(* IEC 61131-3 sources: plc-st-coding-agent/progress/evidence/f14_v3_parallel_20261112/jobs/custom_minimax-m27 (part 3) *)

(* ---- self-hard-02.raw_candidate_01.st ---- *)
FUNCTION_BLOCK FB
VAR_INPUT
    startBtn   : BOOL;
    abortBtn   : BOOL;
    setpoint   : REAL;
    pv         : REAL;
    maxDuration: INT;
END_VAR
VAR_OUTPUT
    elapsed : INT := 0;
    phase   : INT := 0;
    timeout : BOOL := FALSE;
END_VAR
VAR
    prev_startBtn : BOOL := FALSE;
    prev_phase    : INT  := 0;
    risingEdge    : BOOL;
END_VAR

    // Detect rising edge of startBtn before any state changes this scan
    risingEdge := startBtn AND NOT prev_startBtn;

    // Priority 1: abort
    IF abortBtn THEN
        phase   := 9;
        // elapsed and timeout stay frozen (no assignment)

    // Priority 2: new rising edge (only if not aborted this scan)
    ELSIF risingEdge THEN
        elapsed := 0;
        timeout := FALSE;
        phase   := 1;

    // Priority 3: running phases — count and evaluate transition
    ELSIF (prev_phase = 1) OR (prev_phase = 2) THEN
        elapsed := elapsed + 1;

        // Check timeout before setting phase
        IF elapsed >= maxDuration THEN
            timeout := TRUE;
            phase   := 3;
        ELSE
            // Phase transition based on temperature
            IF (prev_phase = 2) OR (pv >= setpoint) THEN
                phase := 2;
            ELSE
                phase := 1;
            END_IF;
        END_IF;

    // Frozen states (phase 0, 3, 9) — no changes to elapsed/phase/timeout
    ELSE
        // phase, elapsed, timeout retain their values
    END_IF;

    // Update previous-cycle snapshot for next scan
    prev_startBtn := startBtn;
    prev_phase    := phase;
END_FUNCTION_BLOCK

(* ---- self-hard-02.raw_candidate_02.st ---- *)
FUNCTION_BLOCK FB
VAR_INPUT
    startBtn   : BOOL;
    abortBtn   : BOOL;
    setpoint   : REAL;
    pv         : REAL;
    maxDuration: INT;
END_VAR
VAR_OUTPUT
    elapsed  : INT  := 0;
    phase    : INT  := 0;
    timeout  : BOOL := FALSE;
END_VAR
VAR
    prev_startBtn : BOOL := FALSE;
    prev_phase    : INT  := 0;
    risingEdge    : BOOL;
END_VAR

    risingEdge := startBtn AND NOT prev_startBtn;

    IF abortBtn THEN
        phase := 9;
        elapsed := elapsed;
        timeout := timeout;

    ELSIF risingEdge THEN
        elapsed := 0;
        timeout := FALSE;
        phase   := 1;

    ELSIF (prev_phase = 1) OR (prev_phase = 2) THEN
        elapsed := elapsed + 1;

        IF elapsed >= maxDuration THEN
            timeout := TRUE;
            phase   := 3;
        ELSE
            IF (prev_phase = 2) OR (pv >= setpoint) THEN
                phase := 2;
            ELSE
                phase := 1;
            END_IF;
        END_IF;

    ELSE
        NULL;
    END_IF;

    prev_startBtn := startBtn;
    prev_phase    := phase;
END_FUNCTION_BLOCK

(* ---- self-hard-03.candidate_01.st ---- *)
FUNCTION_BLOCK FB
VAR_INPUT
    pushEn  : BOOL;
    pushItem: INT;
    popEn   : BOOL;
END_VAR

VAR_INOUT
    fifo : ARRAY[1..8] OF INT;
END_VAR

VAR_OUTPUT
    count : INT;
    full  : BOOL;
    empty : BOOL;
    head  : INT;
END_VAR

VAR
    prevPushEn : BOOL := FALSE;
    prevPopEn  : BOOL := FALSE;
    curCount   : INT  := 0;
    i          : INT;
    risingPush : BOOL;
    risingPop  : BOOL;
END_VAR

(* Detect rising edges *)
risingPush := pushEn AND NOT prevPushEn;
risingPop  := popEn  AND NOT prevPopEn;

(* Update edge memory for next scan *)
prevPushEn := pushEn;
prevPopEn  := popEn;

(* ---- POP (executed first) ---- *)
IF risingPop THEN
    IF curCount > 0 THEN
        (* shift left to remove the oldest element *)
        FOR i := 1 TO curCount - 1 DO
            fifo[i] := fifo[i+1];
        END_FOR;
        curCount := curCount - 1;
    END_IF;
END_IF;

(* ---- PUSH (executed after pop) ---- *)
IF risingPush THEN
    IF curCount < 8 THEN
        curCount := curCount + 1;
        fifo[curCount] := pushItem;
    END_IF;
END_IF;

(* ---- Outputs ---- *)
count := curCount;
full  := (curCount = 8);
empty := (curCount = 0);
head  := IF empty THEN 0 ELSE fifo[1];

END_FUNCTION_BLOCK

(* ---- self-hard-03.candidate_02.st ---- *)
FUNCTION_BLOCK FB
VAR_INPUT
    pushEn  : BOOL;
    pushItem: INT;
    popEn   : BOOL;
END_VAR

VAR_IN_OUT
    fifo : ARRAY[1..8] OF INT;
END_VAR

VAR_OUTPUT
    count : INT;
    full  : BOOL;
    empty : BOOL;
    head  : INT;
END_VAR

VAR
    prevPushEn : BOOL := FALSE;
    prevPopEn  : BOOL := FALSE;
    curCount   : INT  := 0;
    i          : INT;
    risingPush : BOOL;
    risingPop  : BOOL;
END_VAR

risingPush := pushEn AND NOT prevPushEn;
risingPop  := popEn  AND NOT prevPopEn;

prevPushEn := pushEn;
prevPopEn  := popEn;

IF risingPop THEN
    IF curCount > 0 THEN
        FOR i := 1 TO curCount - 1 DO
            fifo[i] := fifo[i+1];
        END_FOR;
        curCount := curCount - 1;
    END_IF;
END_IF;

IF risingPush THEN
    IF curCount < 8 THEN
        curCount := curCount + 1;
        fifo[curCount] := pushItem;
    END_IF;
END_IF;

count := curCount;
full  := (curCount = 8);
empty := (curCount = 0);
head  := fifo[1];

IF empty THEN
    head := 0;
END_IF;

END_FUNCTION_BLOCK

(* ---- self-hard-03.raw_candidate_01.st ---- *)
FUNCTION_BLOCK FB
VAR_INPUT
    pushEn  : BOOL;
    pushItem: INT;
    popEn   : BOOL;
END_VAR

VAR_INOUT
    fifo : ARRAY[1..8] OF INT;
END_VAR

VAR_OUTPUT
    count : INT;
    full  : BOOL;
    empty : BOOL;
    head  : INT;
END_VAR

VAR
    prevPushEn : BOOL := FALSE;
    prevPopEn  : BOOL := FALSE;
    curCount   : INT  := 0;
    i          : INT;
    risingPush : BOOL;
    risingPop  : BOOL;
END_VAR

(* Detect rising edges *)
risingPush := pushEn AND NOT prevPushEn;
risingPop  := popEn  AND NOT prevPopEn;

(* Update edge memory for next scan *)
prevPushEn := pushEn;
prevPopEn  := popEn;

(* ---- POP (executed first) ---- *)
IF risingPop THEN
    IF curCount > 0 THEN
        (* shift left to remove the oldest element *)
        FOR i := 1 TO curCount - 1 DO
            fifo[i] := fifo[i+1];
        END_FOR;
        curCount := curCount - 1;
    END_IF;
END_IF;

(* ---- PUSH (executed after pop) ---- *)
IF risingPush THEN
    IF curCount < 8 THEN
        curCount := curCount + 1;
        fifo[curCount] := pushItem;
    END_IF;
END_IF;

(* ---- Outputs ---- *)
count := curCount;
full  := (curCount = 8);
empty := (curCount = 0);
head  := IF empty THEN 0 ELSE fifo[1];

END_FUNCTION_BLOCK

(* ---- self-hard-03.raw_candidate_02.st ---- *)
FUNCTION_BLOCK FB
VAR_INPUT
    pushEn  : BOOL;
    pushItem: INT;
    popEn   : BOOL;
END_VAR

VAR_IN_OUT
    fifo : ARRAY[1..8] OF INT;
END_VAR

VAR_OUTPUT
    count : INT;
    full  : BOOL;
    empty : BOOL;
    head  : INT;
END_VAR

VAR
    prevPushEn : BOOL := FALSE;
    prevPopEn  : BOOL := FALSE;
    curCount   : INT  := 0;
    i          : INT;
    risingPush : BOOL;
    risingPop  : BOOL;
END_VAR

risingPush := pushEn AND NOT prevPushEn;
risingPop  := popEn  AND NOT prevPopEn;

prevPushEn := pushEn;
prevPopEn  := popEn;

IF risingPop THEN
    IF curCount > 0 THEN
        FOR i := 1 TO curCount - 1 DO
            fifo[i] := fifo[i+1];
        END_FOR;
        curCount := curCount - 1;
    END_IF;
END_IF;

IF risingPush THEN
    IF curCount < 8 THEN
        curCount := curCount + 1;
        fifo[curCount] := pushItem;
    END_IF;
END_IF;

count := curCount;
full  := (curCount = 8);
empty := (curCount = 0);
head  := fifo[1];

IF empty THEN
    head := 0;
END_IF;

END_FUNCTION_BLOCK

(* ---- self-hard-04.candidate_01.st ---- *)
FUNCTION_BLOCK FB
VAR_INPUT
    demand     : INT;
    runHours   : ARRAY[1..5] OF LINT;
    rotated    : BOOL;
END_VAR
VAR_OUTPUT
    leadPump     : INT := 0;
    lagPump      : INT := 0;
    runningCount : INT := 0;
END_VAR
VAR
    prevDemand   : INT  := 0;
    prevLead     : INT  := 0;
    prevLag      : INT  := 0;
    prevRunning  : INT  := 0;
END_VAR

VAR_TEMP
    i            : INT;
    minHours     : LINT;
    minIdx       : INT;
    minHours2    : LINT;
    minIdx2      : INT;
    adjDemand    : INT;
    leadChanged  : BOOL;
    runInc       : BOOL;
END_VAR

// ── 1. 裁剪需求台数 ──────────────────────────────────────────────
IF demand < 0 THEN
    adjDemand := 0;
ELSIF demand > 5 THEN
    adjDemand := 5;
ELSE
    adjDemand := demand;
END_IF;

// ── 2. 需求归零 → 立即清除主备 ───────────────────────────────────
IF adjDemand = 0 THEN
    leadPump     := 0;
    lagPump      := 0;
    runningCount := 0;
    prevDemand   := 0;
    prevLead     := 0;
    prevLag      := 0;
    prevRunning  := 0;
    RETURN;
END_IF;

// ── 3. 主泵选择 ──────────────────────────────────────────────────
// 初选：上次主泵为空（需求从 0 恢复）
IF prevLead = 0 THEN
    minHours := runHours[1];
    minIdx   := 1;
    FOR i := 2 TO 5 DO
        IF runHours[i] < minHours OR (runHours[i] = minHours AND i < minIdx) THEN
            minHours := runHours[i];
            minIdx   := i;
        END_IF;
    END_FOR;
    leadPump := minIdx;
// 轮换请求有效且迟滞条件满足时换主
ELSIF rotated THEN
    // 找全场（工时，泵号）最小者
    minHours := runHours[1];
    minIdx   := 1;
    FOR i := 2 TO 5 DO
        IF runHours[i] < minHours OR (runHours[i] = minHours AND i < minIdx) THEN
            minHours := runHours[i];
            minIdx   := i;
        END_IF;
    END_FOR;
    // 迟滞：本拍主泵工时比最短工时严格多 50h 以上
    IF runHours[prevLead] - minHours > 50 THEN
        leadPump := minIdx;
    ELSE
        leadPump := prevLead;
    END_IF;
ELSE
    // 无请求且有主泵 → 保持
    leadPump := prevLead;
END_IF;

// ── 4. 辅助标记 ──────────────────────────────────────────────────
leadChanged := (leadPump <> prevLead);
runInc      := (adjDemand > prevRunning);

// ── 5. 备泵选择（仅在「初选、换主、运行台数上升」时重选）─────────
IF adjDemand >= 2 THEN
    // 初选：lagPump 仍为 0
    // 换主或台数上升：lagPump 需要刷新
    IF lagPump = 0 OR leadChanged OR runInc THEN
        // 找除主泵外（工时，泵号）最小者
        minHours2 := LINT#16#7FFFFFFFFFFFFFFF;  // 最大值
        minIdx2   := 0;
        FOR i := 1 TO 5 DO
            IF i <> leadPump THEN
                IF runHours[i] < minHours2 OR (runHours[i] = minHours2 AND i < minIdx2) THEN
                    minHours2 := runHours[i];
                    minIdx2   := i;
                END_IF;
            END_IF;
        END_FOR;
        lagPump := minIdx2;
    ELSE
        // 主泵未变且台数未升 → 保持原备泵（S9 约束）
        lagPump := prevLag;
    END_IF;
ELSE
    // 需求 1 台 → 无备泵
    lagPump := 0;
END_IF;

// ── 6. 运行台数 & 状态快照 ───────────────────────────────────────
runningCount := adjDemand;
prevDemand   := adjDemand;
prevLead     := leadPump;
prevLag      := lagPump;
prevRunning  := runningCount;
END_FUNCTION_BLOCK

(* ---- self-hard-04.candidate_02.st ---- *)
FUNCTION_BLOCK FB
VAR_INPUT
    demand   : INT;
    runHours : ARRAY[1..5] OF LINT;
    rotated  : BOOL;
END_VAR
VAR_OUTPUT
    leadPump     : INT := 0;
    lagPump      : INT := 0;
    runningCount : INT := 0;
END_VAR
VAR
    prevDemand     : INT  := -1;
    prevLead       : INT  := 0;
    prevLag        : INT  := 0;
    prevRunning    : INT  := 0;
    firstPositive  : BOOL := FALSE;
END_VAR
VAR_TEMP
    i           : INT;
    minHours    : LINT;
    minIdx      : INT;
    minHours2   : LINT;
    minIdx2     : INT;
    adjDemand   : INT;
    leadChanged : BOOL;
    runInc      : BOOL;
END_VAR

// ── 裁剪需求台数 ──────────────────────────────────────────────────
IF demand < 0 THEN
    adjDemand := 0;
ELSIF demand > 5 THEN
    adjDemand := 5;
ELSE
    adjDemand := demand;
END_IF;

// ── 首次调用：初始化 prevDemand ──────────────────────────────────
IF prevDemand = -1 THEN
    prevDemand := adjDemand;
END_IF;

// ── 需求为 0：清空主备 ───────────────────────────────────────────
IF adjDemand = 0 THEN
    leadPump     := 0;
    lagPump      := 0;
    runningCount := 0;
    prevLead     := 0;
    prevLag      := 0;
    prevRunning  := 0;
    firstPositive := FALSE;
    prevDemand    := 0;
    RETURN;
END_IF;

// ── 主泵选择 ──────────────────────────────────────────────────────
// 初始选择：首次正需求
IF firstPositive THEN
    minHours := runHours[1];
    minIdx   := 1;
    FOR i := 2 TO 5 DO
        IF runHours[i] < minHours OR (runHours[i] = minHours AND i < minIdx) THEN
            minHours := runHours[i];
            minIdx   := i;
        END_IF;
    END_FOR;
    leadPump := minIdx;
// 迟滞换主：轮换请求有效 且 原主泵工时比全场最短严格多 50h 以上
ELSIF rotated AND prevLead <> 0 THEN
    minHours := runHours[1];
    minIdx   := 1;
    FOR i := 2 TO 5 DO
        IF runHours[i] < minHours OR (runHours[i] = minHours AND i < minIdx) THEN
            minHours := runHours[i];
            minIdx   := i;
        END_IF;
    END_FOR;
    IF runHours[prevLead] - minHours > 50 THEN
        leadPump := minIdx;
    ELSE
        leadPump := prevLead;
    END_IF;
ELSE
    leadPump := prevLead;
END_IF;

// ── 辅助标记 ──────────────────────────────────────────────────────
leadChanged := (leadPump <> prevLead);
runInc      := (adjDemand > prevRunning);

// ── 备泵选择（仅「初选、换主、运行台数上升」时重选）──────────────
IF adjDemand >= 2 THEN
    IF lagPump = 0 OR leadChanged OR runInc THEN
        minHours2 := LINT#16#7FFFFFFFFFFFFFFF;
        minIdx2   := 0;
        FOR i := 1 TO 5 DO
            IF i <> leadPump THEN
                IF runHours[i] < minHours2 OR (runHours[i] = minHours2 AND i < minIdx2) THEN
                    minHours2 := runHours[i];
                    minIdx2   := i;
                END_IF;
            END_IF;
        END_FOR;
        lagPump := minIdx2;
    ELSE
        lagPump := prevLag;
    END_IF;
ELSE
    lagPump := 0;
END_IF;

// ── 运行台数 & 状态快照 ──────────────────────────────────────────
runningCount  := adjDemand;
firstPositive := FALSE;
prevLead      := leadPump;
prevLag       := lagPump;
prevRunning   := runningCount;
prevDemand    := adjDemand;
END_FUNCTION_BLOCK

(* ---- self-hard-04.raw_candidate_01.st ---- *)
FUNCTION_BLOCK FB
VAR_INPUT
    demand     : INT;
    runHours   : ARRAY[1..5] OF LINT;
    rotated    : BOOL;
END_VAR
VAR_OUTPUT
    leadPump     : INT := 0;
    lagPump      : INT := 0;
    runningCount : INT := 0;
END_VAR
VAR
    prevDemand   : INT  := 0;
    prevLead     : INT  := 0;
    prevLag      : INT  := 0;
    prevRunning  : INT  := 0;
END_VAR

VAR_TEMP
    i            : INT;
    minHours     : LINT;
    minIdx       : INT;
    minHours2    : LINT;
    minIdx2      : INT;
    adjDemand    : INT;
    leadChanged  : BOOL;
    runInc       : BOOL;
END_VAR

// ── 1. 裁剪需求台数 ──────────────────────────────────────────────
IF demand < 0 THEN
    adjDemand := 0;
ELSIF demand > 5 THEN
    adjDemand := 5;
ELSE
    adjDemand := demand;
END_IF;

// ── 2. 需求归零 → 立即清除主备 ───────────────────────────────────
IF adjDemand = 0 THEN
    leadPump     := 0;
    lagPump      := 0;
    runningCount := 0;
    prevDemand   := 0;
    prevLead     := 0;
    prevLag      := 0;
    prevRunning  := 0;
    RETURN;
END_IF;

// ── 3. 主泵选择 ──────────────────────────────────────────────────
// 初选：上次主泵为空（需求从 0 恢复）
IF prevLead = 0 THEN
    minHours := runHours[1];
    minIdx   := 1;
    FOR i := 2 TO 5 DO
        IF runHours[i] < minHours OR (runHours[i] = minHours AND i < minIdx) THEN
            minHours := runHours[i];
            minIdx   := i;
        END_IF;
    END_FOR;
    leadPump := minIdx;
// 轮换请求有效且迟滞条件满足时换主
ELSIF rotated THEN
    // 找全场（工时，泵号）最小者
    minHours := runHours[1];
    minIdx   := 1;
    FOR i := 2 TO 5 DO
        IF runHours[i] < minHours OR (runHours[i] = minHours AND i < minIdx) THEN
            minHours := runHours[i];
            minIdx   := i;
        END_IF;
    END_FOR;
    // 迟滞：本拍主泵工时比最短工时严格多 50h 以上
    IF runHours[prevLead] - minHours > 50 THEN
        leadPump := minIdx;
    ELSE
        leadPump := prevLead;
    END_IF;
ELSE
    // 无请求且有主泵 → 保持
    leadPump := prevLead;
END_IF;

// ── 4. 辅助标记 ──────────────────────────────────────────────────
leadChanged := (leadPump <> prevLead);
runInc      := (adjDemand > prevRunning);

// ── 5. 备泵选择（仅在「初选、换主、运行台数上升」时重选）─────────
IF adjDemand >= 2 THEN
    // 初选：lagPump 仍为 0
    // 换主或台数上升：lagPump 需要刷新
    IF lagPump = 0 OR leadChanged OR runInc THEN
        // 找除主泵外（工时，泵号）最小者
        minHours2 := LINT#16#7FFFFFFFFFFFFFFF;  // 最大值
        minIdx2   := 0;
        FOR i := 1 TO 5 DO
            IF i <> leadPump THEN
                IF runHours[i] < minHours2 OR (runHours[i] = minHours2 AND i < minIdx2) THEN
                    minHours2 := runHours[i];
                    minIdx2   := i;
                END_IF;
            END_IF;
        END_FOR;
        lagPump := minIdx2;
    ELSE
        // 主泵未变且台数未升 → 保持原备泵（S9 约束）
        lagPump := prevLag;
    END_IF;
ELSE
    // 需求 1 台 → 无备泵
    lagPump := 0;
END_IF;

// ── 6. 运行台数 & 状态快照 ───────────────────────────────────────
runningCount := adjDemand;
prevDemand   := adjDemand;
prevLead     := leadPump;
prevLag      := lagPump;
prevRunning  := runningCount;
END_FUNCTION_BLOCK

(* ---- self-hard-04.raw_candidate_02.st ---- *)
FUNCTION_BLOCK FB
VAR_INPUT
    demand   : INT;
    runHours : ARRAY[1..5] OF LINT;
    rotated  : BOOL;
END_VAR
VAR_OUTPUT
    leadPump     : INT := 0;
    lagPump      : INT := 0;
    runningCount : INT := 0;
END_VAR
VAR
    prevDemand     : INT  := -1;
    prevLead       : INT  := 0;
    prevLag        : INT  := 0;
    prevRunning    : INT  := 0;
    firstPositive  : BOOL := FALSE;
END_VAR
VAR_TEMP
    i           : INT;
    minHours    : LINT;
    minIdx      : INT;
    minHours2   : LINT;
    minIdx2     : INT;
    adjDemand   : INT;
    leadChanged : BOOL;
    runInc      : BOOL;
END_VAR

// ── 裁剪需求台数 ──────────────────────────────────────────────────
IF demand < 0 THEN
    adjDemand := 0;
ELSIF demand > 5 THEN
    adjDemand := 5;
ELSE
    adjDemand := demand;
END_IF;

// ── 首次调用：初始化 prevDemand ──────────────────────────────────
IF prevDemand = -1 THEN
    prevDemand := adjDemand;
END_IF;

// ── 需求为 0：清空主备 ───────────────────────────────────────────
IF adjDemand = 0 THEN
    leadPump     := 0;
    lagPump      := 0;
    runningCount := 0;
    prevLead     := 0;
    prevLag      := 0;
    prevRunning  := 0;
    firstPositive := FALSE;
    prevDemand    := 0;
    RETURN;
END_IF;

// ── 主泵选择 ──────────────────────────────────────────────────────
// 初始选择：首次正需求
IF firstPositive THEN
    minHours := runHours[1];
    minIdx   := 1;
    FOR i := 2 TO 5 DO
        IF runHours[i] < minHours OR (runHours[i] = minHours AND i < minIdx) THEN
            minHours := runHours[i];
            minIdx   := i;
        END_IF;
    END_FOR;
    leadPump := minIdx;
// 迟滞换主：轮换请求有效 且 原主泵工时比全场最短严格多 50h 以上
ELSIF rotated AND prevLead <> 0 THEN
    minHours := runHours[1];
    minIdx   := 1;
    FOR i := 2 TO 5 DO
        IF runHours[i] < minHours OR (runHours[i] = minHours AND i < minIdx) THEN
            minHours := runHours[i];
            minIdx   := i;
        END_IF;
    END_FOR;
    IF runHours[prevLead] - minHours > 50 THEN
        leadPump := minIdx;
    ELSE
        leadPump := prevLead;
    END_IF;
ELSE
    leadPump := prevLead;
END_IF;

// ── 辅助标记 ──────────────────────────────────────────────────────
leadChanged := (leadPump <> prevLead);
runInc      := (adjDemand > prevRunning);

// ── 备泵选择（仅「初选、换主、运行台数上升」时重选）──────────────
IF adjDemand >= 2 THEN
    IF lagPump = 0 OR leadChanged OR runInc THEN
        minHours2 := LINT#16#7FFFFFFFFFFFFFFF;
        minIdx2   := 0;
        FOR i := 1 TO 5 DO
            IF i <> leadPump THEN
                IF runHours[i] < minHours2 OR (runHours[i] = minHours2 AND i < minIdx2) THEN
                    minHours2 := runHours[i];
                    minIdx2   := i;
                END_IF;
            END_IF;
        END_FOR;
        lagPump := minIdx2;
    ELSE
        lagPump := prevLag;
    END_IF;
ELSE
    lagPump := 0;
END_IF;

// ── 运行台数 & 状态快照 ──────────────────────────────────────────
runningCount  := adjDemand;
firstPositive := FALSE;
prevLead      := leadPump;
prevLag       := lagPump;
prevRunning   := runningCount;
prevDemand    := adjDemand;
END_FUNCTION_BLOCK

(* ---- self-hard-05.candidate_01.st ---- *)
FUNCTION_BLOCK FB
VAR_INPUT
    runRequest  : BOOL;
    flameOK     : BOOL;
    o2Valid     : BOOL;
    o2PV        : REAL;
    baseAir     : REAL;
    resetBtn    : BOOL;
END_VAR
VAR_OUTPUT
    fuelPermit  : BOOL;
    trimEnable  : BOOL;
    airTrim     : REAL;
    airCommand  : REAL;
    tripLatched : BOOL;
    o2Fault     : BOOL;
END_VAR
VAR
    prevResetBtn : BOOL := FALSE;
END_VAR

    // Rising edge detection for reset button
    VAR
        resetRisingEdge : BOOL;
    END_VAR
    resetRisingEdge := resetBtn AND NOT prevResetBtn;
    prevResetBtn := resetBtn;

    // Trip latch: immediate set on flame loss during run; clear only on safe-state reset edge
    IF runRequest AND NOT flameOK THEN
        tripLatched := TRUE;
    ELSIF resetRisingEdge AND NOT runRequest AND NOT flameOK THEN
        tripLatched := FALSE;
    END_IF;

    // Fuel permit
    fuelPermit := runRequest AND flameOK AND NOT tripLatched;

    // O2 analyzer fault
    o2Fault := NOT o2Valid OR o2PV < 0.0 OR o2PV > 21.0;

    // Trim enable
    trimEnable := fuelPermit AND NOT o2Fault;

    // Air trim: compute and clamp to [-10, +10]; force 0 when trim not enabled
    IF trimEnable THEN
        airTrim := 2.0 * (2.0 - o2PV);
        IF airTrim > 10.0 THEN
            airTrim := 10.0;
        ELSIF airTrim < -10.0 THEN
            airTrim := -10.0;
        END_IF;
    ELSE
        airTrim := 0.0;
    END_IF;

    // Air command: sum and clamp to [0, 100]; force 0 when no fuel permit
    IF fuelPermit THEN
        airCommand := baseAir + airTrim;
        IF airCommand > 100.0 THEN
            airCommand := 100.0;
        ELSIF airCommand < 0.0 THEN
            airCommand := 0.0;
        END_IF;
    ELSE
        airCommand := 0.0;
    END_IF;
END_FUNCTION_BLOCK

(* ---- self-hard-05.raw_candidate_01.st ---- *)
FUNCTION_BLOCK FB
VAR_INPUT
    runRequest  : BOOL;
    flameOK     : BOOL;
    o2Valid     : BOOL;
    o2PV        : REAL;
    baseAir     : REAL;
    resetBtn    : BOOL;
END_VAR
VAR_OUTPUT
    fuelPermit  : BOOL;
    trimEnable  : BOOL;
    airTrim     : REAL;
    airCommand  : REAL;
    tripLatched : BOOL;
    o2Fault     : BOOL;
END_VAR
VAR
    prevResetBtn : BOOL := FALSE;
END_VAR

    // Rising edge detection for reset button
    VAR
        resetRisingEdge : BOOL;
    END_VAR
    resetRisingEdge := resetBtn AND NOT prevResetBtn;
    prevResetBtn := resetBtn;

    // Trip latch: immediate set on flame loss during run; clear only on safe-state reset edge
    IF runRequest AND NOT flameOK THEN
        tripLatched := TRUE;
    ELSIF resetRisingEdge AND NOT runRequest AND NOT flameOK THEN
        tripLatched := FALSE;
    END_IF;

    // Fuel permit
    fuelPermit := runRequest AND flameOK AND NOT tripLatched;

    // O2 analyzer fault
    o2Fault := NOT o2Valid OR o2PV < 0.0 OR o2PV > 21.0;

    // Trim enable
    trimEnable := fuelPermit AND NOT o2Fault;

    // Air trim: compute and clamp to [-10, +10]; force 0 when trim not enabled
    IF trimEnable THEN
        airTrim := 2.0 * (2.0 - o2PV);
        IF airTrim > 10.0 THEN
            airTrim := 10.0;
        ELSIF airTrim < -10.0 THEN
            airTrim := -10.0;
        END_IF;
    ELSE
        airTrim := 0.0;
    END_IF;

    // Air command: sum and clamp to [0, 100]; force 0 when no fuel permit
    IF fuelPermit THEN
        airCommand := baseAir + airTrim;
        IF airCommand > 100.0 THEN
            airCommand := 100.0;
        ELSIF airCommand < 0.0 THEN
            airCommand := 0.0;
        END_IF;
    ELSE
        airCommand := 0.0;
    END_IF;
END_FUNCTION_BLOCK

(* ---- self-hard-06.candidate_01.st ---- *)
TYPE ETripStickingState :
(
   ST_CLEAR := 0,
   ST_COUNT1 := 1,
   ST_COUNT2 := 2,
   ST_CONFIRMED := 3
);
END_TYPE;

FUNCTION_BLOCK FB
VAR_INPUT
    runRequest       : BOOL;
    pressure         : REAL;
    pressureValid    : BOOL;
    fuelFlow         : REAL;
    steamFlow        : REAL;
    outletCmd        : INT;
    outletFeedback   : INT;
    resetBtn         : BOOL;
END_VAR
VAR_OUTPUT
    tripLatched      : BOOL;
    fuelPermit       : BOOL;
    currentCauseMask : WORD;
    latchedCauseMask : WORD;
    diagnosticActive : BOOL;
END_VAR
VAR
    prevCondSticking : BOOL := FALSE;
    stickingCounter  : UINT  := 0;
    prevResetBtn     : BOOL  := FALSE;
END_VAR
VAR_CONSTANT
    cPressureTrip     : REAL := 4500.0;
    cPressureReset    : REAL := 4200.0;
    cFuelFlowThreshold: REAL := 4.0;
    cSteamFlowThreshold: REAL := 10.0;
    cStickingCycles   : UINT := 3;
    cValveCmdMin      : INT  := 50;
    cValveFbkMax      : INT  := 10;
END_VAR
VAR_TEMP
    risingEdgeReset : BOOL;
    validReset      : BOOL;
    tripCondition   : BOOL;
    condSticking    : BOOL;
    bit0            : BOOL;
    bit1            : BOOL;
    bit2            : BOOL;
    bit3            : BOOL;
END_VAR

    risingEdgeReset := resetBtn AND NOT prevResetBtn;

    validReset := risingEdgeReset
                  AND NOT runRequest
                  AND pressureValid
                  AND (pressure <= cPressureReset);

    IF validReset THEN
        tripLatched      := FALSE;
        latchedCauseMask := 0;
    ELSE
        tripCondition := runRequest AND (NOT pressureValid OR pressure >= cPressureTrip);
        IF tripCondition THEN
            tripLatched := TRUE;
        END_IF;
        IF tripLatched THEN
            latchedCauseMask := latchedCauseMask OR currentCauseMask;
        END_IF;
    END_IF;

    fuelPermit := runRequest AND NOT tripLatched;

    condSticking := runRequest
                    AND pressureValid
                    AND (pressure >= cPressureTrip)
                    AND (outletCmd >= cValveCmdMin)
                    AND (outletFeedback <= cValveFbkMax);

    IF condSticking THEN
        IF stickingCounter < cStickingCycles THEN
            stickingCounter := stickingCounter + 1;
        END_IF;
    ELSE
        stickingCounter := 0;
    END_IF;

    prevCondSticking := condSticking;

    IF NOT runRequest THEN
        currentCauseMask := 0;
    ELSIF NOT pressureValid THEN
        currentCauseMask := 1;
    ELSIF pressure >= cPressureTrip THEN
        bit0 := FALSE;
        bit1 := (stickingCounter >= cStickingCycles)
                AND prevCondSticking;
        bit2 := (fuelFlow >= cFuelFlowThreshold)
                AND (steamFlow <= cSteamFlowThreshold);
        bit3 := NOT bit1 AND NOT bit2;
        currentCauseMask := TO_WORD(
            TO_INT(bit0) +
            TO_INT(bit1) * 2 +
            TO_INT(bit2) * 4 +
            TO_INT(bit3) * 8
        );
    ELSE
        currentCauseMask := 0;
    END_IF;

    diagnosticActive := (currentCauseMask <> 0);

    prevResetBtn := resetBtn;
END_FUNCTION_BLOCK

(* ---- self-hard-06.candidate_02.st ---- *)
TYPE ETripStickingState :
(
   ST_CLEAR := 0,
   ST_COUNT1 := 1,
   ST_COUNT2 := 2,
   ST_CONFIRMED := 3
);
END_TYPE;

FUNCTION_BLOCK FB
VAR_INPUT
    runRequest       : BOOL;
    pressure         : REAL;
    pressureValid    : BOOL;
    fuelFlow         : REAL;
    steamFlow        : REAL;
    outletCmd        : INT;
    outletFeedback   : INT;
    resetBtn         : BOOL;
END_VAR
VAR_OUTPUT
    tripLatched      : BOOL;
    fuelPermit       : BOOL;
    currentCauseMask : WORD;
    latchedCauseMask : WORD;
    diagnosticActive : BOOL;
END_VAR
VAR
    prevCondSticking : BOOL := FALSE;
    stickingCounter  : UINT := 0;
    prevResetBtn     : BOOL := FALSE;
END_VAR
VAR_TEMP
    risingEdgeReset : BOOL;
    validReset      : BOOL;
    tripCondition   : BOOL;
    condSticking    : BOOL;
    stuckConfirmed  : BOOL;
    bit2            : BOOL;
END_VAR

    risingEdgeReset := resetBtn AND NOT prevResetBtn;

    validReset := risingEdgeReset
                  AND (NOT runRequest)
                  AND pressureValid
                  AND (pressure <= 4200.0);

    IF validReset THEN
        tripLatched      := FALSE;
        latchedCauseMask := 0;
    ELSE
        tripCondition := runRequest AND (NOT pressureValid OR pressure >= 4500.0);
        IF tripCondition THEN
            tripLatched := TRUE;
        END_IF;
        IF tripLatched THEN
            latchedCauseMask := latchedCauseMask OR currentCauseMask;
        END_IF;
    END_IF;

    fuelPermit := runRequest AND NOT tripLatched;

    condSticking := runRequest
                    AND pressureValid
                    AND (pressure >= 4500.0)
                    AND (outletCmd >= 50)
                    AND (outletFeedback <= 10);

    IF condSticking THEN
        IF stickingCounter < 16#FFFF THEN
            stickingCounter := stickingCounter + 1;
        END_IF;
    ELSE
        stickingCounter := 0;
    END_IF;

    stuckConfirmed := (stickingCounter >= 3) AND prevCondSticking;

    bit2 := (fuelFlow >= 4.0) AND (steamFlow <= 10.0);

    IF NOT runRequest THEN
        currentCauseMask := 0;
    ELSIF NOT pressureValid THEN
        currentCauseMask := 1;
    ELSIF pressure >= 4500.0 THEN
        currentCauseMask := TO_WORD(
            TO_INT(stuckConfirmed) * 2 +
            TO_INT(bit2) * 4 +
            TO_INT(NOT stuckConfirmed AND NOT bit2) * 8
        );
    ELSE
        currentCauseMask := 0;
    END_IF;

    diagnosticActive := (currentCauseMask <> 0);

    prevCondSticking := condSticking;
    prevResetBtn     := resetBtn;
END_FUNCTION_BLOCK

(* ---- self-hard-06.raw_candidate_01.st ---- *)
TYPE ETripStickingState :
(
   ST_CLEAR := 0,
   ST_COUNT1 := 1,
   ST_COUNT2 := 2,
   ST_CONFIRMED := 3
);
END_TYPE

FUNCTION_BLOCK FB
VAR_INPUT
    runRequest       : BOOL;
    pressure         : REAL;
    pressureValid    : BOOL;
    fuelFlow         : REAL;
    steamFlow        : REAL;
    outletCmd        : INT;
    outletFeedback   : INT;
    resetBtn         : BOOL;
END_VAR
VAR_OUTPUT
    tripLatched      : BOOL;
    fuelPermit       : BOOL;
    currentCauseMask : WORD;
    latchedCauseMask : WORD;
    diagnosticActive : BOOL;
END_VAR
VAR
    prevCondSticking : BOOL := FALSE;
    stickingCounter  : UINT  := 0;
    prevResetBtn     : BOOL  := FALSE;
END_VAR
VAR_CONSTANT
    cPressureTrip     : REAL := 4500.0;
    cPressureReset    : REAL := 4200.0;
    cFuelFlowThreshold: REAL := 4.0;
    cSteamFlowThreshold: REAL := 10.0;
    cStickingCycles   : UINT := 3;
    cValveCmdMin      : INT  := 50;
    cValveFbkMax      : INT  := 10;
END_VAR
VAR_TEMP
    risingEdgeReset : BOOL;
    validReset      : BOOL;
    tripCondition   : BOOL;
    condSticking    : BOOL;
    bit0            : BOOL;
    bit1            : BOOL;
    bit2            : BOOL;
    bit3            : BOOL;
END_VAR

    risingEdgeReset := resetBtn AND NOT prevResetBtn;

    validReset := risingEdgeReset
                  AND NOT runRequest
                  AND pressureValid
                  AND (pressure <= cPressureReset);

    IF validReset THEN
        tripLatched      := FALSE;
        latchedCauseMask := 0;
    ELSE
        tripCondition := runRequest AND (NOT pressureValid OR pressure >= cPressureTrip);
        IF tripCondition THEN
            tripLatched := TRUE;
        END_IF;
        IF tripLatched THEN
            latchedCauseMask := latchedCauseMask OR currentCauseMask;
        END_IF;
    END_IF;

    fuelPermit := runRequest AND NOT tripLatched;

    condSticking := runRequest
                    AND pressureValid
                    AND (pressure >= cPressureTrip)
                    AND (outletCmd >= cValveCmdMin)
                    AND (outletFeedback <= cValveFbkMax);

    IF condSticking THEN
        IF stickingCounter < cStickingCycles THEN
            stickingCounter := stickingCounter + 1;
        END_IF;
    ELSE
        stickingCounter := 0;
    END_IF;

    prevCondSticking := condSticking;

    IF NOT runRequest THEN
        currentCauseMask := 0;
    ELSIF NOT pressureValid THEN
        currentCauseMask := 1;
    ELSIF pressure >= cPressureTrip THEN
        bit0 := FALSE;
        bit1 := (stickingCounter >= cStickingCycles)
                AND prevCondSticking;
        bit2 := (fuelFlow >= cFuelFlowThreshold)
                AND (steamFlow <= cSteamFlowThreshold);
        bit3 := NOT bit1 AND NOT bit2;
        currentCauseMask := TO_WORD(
            TO_INT(bit0) +
            TO_INT(bit1) * 2 +
            TO_INT(bit2) * 4 +
            TO_INT(bit3) * 8
        );
    ELSE
        currentCauseMask := 0;
    END_IF;

    diagnosticActive := (currentCauseMask <> 0);

    prevResetBtn := resetBtn;
END_FUNCTION_BLOCK

(* ---- self-hard-06.raw_candidate_02.st ---- *)
TYPE ETripStickingState :
(
   ST_CLEAR := 0,
   ST_COUNT1 := 1,
   ST_COUNT2 := 2,
   ST_CONFIRMED := 3
);
END_TYPE;

FUNCTION_BLOCK FB
VAR_INPUT
    runRequest       : BOOL;
    pressure         : REAL;
    pressureValid    : BOOL;
    fuelFlow         : REAL;
    steamFlow        : REAL;
    outletCmd        : INT;
    outletFeedback   : INT;
    resetBtn         : BOOL;
END_VAR
VAR_OUTPUT
    tripLatched      : BOOL;
    fuelPermit       : BOOL;
    currentCauseMask : WORD;
    latchedCauseMask : WORD;
    diagnosticActive : BOOL;
END_VAR
VAR
    prevCondSticking : BOOL := FALSE;
    stickingCounter  : UINT := 0;
    prevResetBtn     : BOOL := FALSE;
END_VAR
VAR_TEMP
    risingEdgeReset : BOOL;
    validReset      : BOOL;
    tripCondition   : BOOL;
    condSticking    : BOOL;
    stuckConfirmed  : BOOL;
    bit2            : BOOL;
END_VAR

    risingEdgeReset := resetBtn AND NOT prevResetBtn;

    validReset := risingEdgeReset
                  AND (NOT runRequest)
                  AND pressureValid
                  AND (pressure <= 4200.0);

    IF validReset THEN
        tripLatched      := FALSE;
        latchedCauseMask := 0;
    ELSE
        tripCondition := runRequest AND (NOT pressureValid OR pressure >= 4500.0);
        IF tripCondition THEN
            tripLatched := TRUE;
        END_IF;
        IF tripLatched THEN
            latchedCauseMask := latchedCauseMask OR currentCauseMask;
        END_IF;
    END_IF;

    fuelPermit := runRequest AND NOT tripLatched;

    condSticking := runRequest
                    AND pressureValid
                    AND (pressure >= 4500.0)
                    AND (outletCmd >= 50)
                    AND (outletFeedback <= 10);

    IF condSticking THEN
        IF stickingCounter < 16#FFFF THEN
            stickingCounter := stickingCounter + 1;
        END_IF;
    ELSE
        stickingCounter := 0;
    END_IF;

    stuckConfirmed := (stickingCounter >= 3) AND prevCondSticking;

    bit2 := (fuelFlow >= 4.0) AND (steamFlow <= 10.0);

    IF NOT runRequest THEN
        currentCauseMask := 0;
    ELSIF NOT pressureValid THEN
        currentCauseMask := 1;
    ELSIF pressure >= 4500.0 THEN
        currentCauseMask := TO_WORD(
            TO_INT(stuckConfirmed) * 2 +
            TO_INT(bit2) * 4 +
            TO_INT(NOT stuckConfirmed AND NOT bit2) * 8
        );
    ELSE
        currentCauseMask := 0;
    END_IF;

    diagnosticActive := (currentCauseMask <> 0);

    prevCondSticking := condSticking;
    prevResetBtn     := resetBtn;
END_FUNCTION_BLOCK

(* ---- self-hard-07.candidate_01.st ---- *)
FUNCTION_BLOCK FB
VAR_INPUT
    mode            : INT;
    resetBtn        : BOOL;
    scanSeconds     : REAL;
    tempSP          : REAL;
    tempPV          : REAL;
    flowPV          : REAL;
    manualFlowSP    : REAL;
    manualValve     : REAL;
END_VAR
VAR_OUTPUT
    flowSP          : REAL;
    valveCommand    : REAL;
    fault           : BOOL;
    normalMode      : BOOL;
END_VAR
VAR
    prevMode        : INT;
    prevFlowSP      : REAL;
    prevValveCommand: REAL;
    prevResetBtn    : BOOL;
    firstScanDone   : BOOL;
    accT            : REAL;
    accF            : REAL;
END_VAR

VAR_TEMP
    isResetRising   : BOOL;
    isModeChange    : BOOL;
    eT              : REAL;
    eF              : REAL;
    trialT          : REAL;
    trialF          : REAL;
    flowSPLimit     : REAL;
    valveLimit      : REAL;
END_VAR

    isResetRising := resetBtn AND NOT prevResetBtn;
    isModeChange := firstScanDone AND (mode <> prevMode);

    fault := (mode < 0) OR (mode > 2) OR (scanSeconds <= 0.0) OR (scanSeconds > 10.0);

    IF isResetRising THEN
        flowSP := manualFlowSP;
        valveCommand := manualValve;
        accT := manualFlowSP - 1.0 * (tempSP - tempPV);
        accF := manualValve - 2.0 * (manualFlowSP - flowPV);
        normalMode := FALSE;
    ELSIF NOT firstScanDone THEN
        flowSP := manualFlowSP;
        valveCommand := manualValve;
        accT := manualFlowSP - 1.0 * (tempSP - tempPV);
        accF := manualValve - 2.0 * (manualFlowSP - flowPV);
        normalMode := FALSE;
    ELSIF fault THEN
        flowSP := manualFlowSP;
        valveCommand := manualValve;
        accT := manualFlowSP - 1.0 * (tempSP - tempPV);
        accF := manualValve - 2.0 * (manualFlowSP - flowPV);
        normalMode := FALSE;
    ELSIF isModeChange THEN
        IF mode = 2 THEN
            flowSP := prevFlowSP;
            valveCommand := prevValveCommand;
            eT := tempSP - tempPV;
            accT := flowSP - 1.0 * eT;
            eF := flowSP - flowPV;
            accF := valveCommand - 2.0 * eF;
        ELSE
            flowSP := manualFlowSP;
            valveCommand := prevValveCommand;
            eT := tempSP - tempPV;
            accT := flowSP - 1.0 * eT;
            eF := flowSP - flowPV;
            accF := valveCommand - 2.0 * eF;
        END_IF;
        normalMode := FALSE;
    ELSE
        normalMode := TRUE;
        eT := tempSP - tempPV;
        eF := flowSP - flowPV;
        IF mode = 2 THEN
            trialT := accT + 0.2 * eT * scanSeconds;
            flowSPLimit := LIMIT(0.0, 1.0 * eT + trialT, 50.0);
            flowSP := flowSPLimit;
            accT := flowSP - 1.0 * eT;
            eF := flowSP - flowPV;
            trialF := accF + 0.5 * eF * scanSeconds;
            valveLimit := LIMIT(0.0, 2.0 * eF + trialF, 100.0);
            valveCommand := valveLimit;
            accF := valveCommand - 2.0 * eF;
        ELSIF mode = 1 THEN
            flowSP := manualFlowSP;
            eF := flowSP - flowPV;
            trialF := accF + 0.5 * eF * scanSeconds;
            valveLimit := LIMIT(0.0, 2.0 * eF + trialF, 100.0);
            valveCommand := valveLimit;
            accF := valveCommand - 2.0 * eF;
        ELSE
            flowSP := manualFlowSP;
            valveCommand := manualValve;
            accF := valveCommand - 2.0 * eF;
        END_IF;
    END_IF;

    prevResetBtn := resetBtn;
    prevMode := mode;
    prevFlowSP := flowSP;
    prevValveCommand := valveCommand;
    firstScanDone := TRUE;
END_FUNCTION_BLOCK

(* ---- self-hard-07.raw_candidate_01.st ---- *)
FUNCTION_BLOCK FB
VAR_INPUT
    mode            : INT;
    resetBtn        : BOOL;
    scanSeconds     : REAL;
    tempSP          : REAL;
    tempPV          : REAL;
    flowPV          : REAL;
    manualFlowSP    : REAL;
    manualValve     : REAL;
END_VAR
VAR_OUTPUT
    flowSP          : REAL;
    valveCommand    : REAL;
    fault           : BOOL;
    normalMode      : BOOL;
END_VAR
VAR
    prevMode        : INT;
    prevFlowSP      : REAL;
    prevValveCommand: REAL;
    prevResetBtn    : BOOL;
    firstScanDone   : BOOL;
    accT            : REAL;
    accF            : REAL;
END_VAR

VAR_TEMP
    isResetRising   : BOOL;
    isModeChange    : BOOL;
    eT              : REAL;
    eF              : REAL;
    trialT          : REAL;
    trialF          : REAL;
    flowSPLimit     : REAL;
    valveLimit      : REAL;
END_VAR

    isResetRising := resetBtn AND NOT prevResetBtn;
    isModeChange := firstScanDone AND (mode <> prevMode);

    fault := (mode < 0) OR (mode > 2) OR (scanSeconds <= 0.0) OR (scanSeconds > 10.0);

    IF isResetRising THEN
        flowSP := manualFlowSP;
        valveCommand := manualValve;
        accT := manualFlowSP - 1.0 * (tempSP - tempPV);
        accF := manualValve - 2.0 * (manualFlowSP - flowPV);
        normalMode := FALSE;
    ELSIF NOT firstScanDone THEN
        flowSP := manualFlowSP;
        valveCommand := manualValve;
        accT := manualFlowSP - 1.0 * (tempSP - tempPV);
        accF := manualValve - 2.0 * (manualFlowSP - flowPV);
        normalMode := FALSE;
    ELSIF fault THEN
        flowSP := manualFlowSP;
        valveCommand := manualValve;
        accT := manualFlowSP - 1.0 * (tempSP - tempPV);
        accF := manualValve - 2.0 * (manualFlowSP - flowPV);
        normalMode := FALSE;
    ELSIF isModeChange THEN
        IF mode = 2 THEN
            flowSP := prevFlowSP;
            valveCommand := prevValveCommand;
            eT := tempSP - tempPV;
            accT := flowSP - 1.0 * eT;
            eF := flowSP - flowPV;
            accF := valveCommand - 2.0 * eF;
        ELSE
            flowSP := manualFlowSP;
            valveCommand := prevValveCommand;
            eT := tempSP - tempPV;
            accT := flowSP - 1.0 * eT;
            eF := flowSP - flowPV;
            accF := valveCommand - 2.0 * eF;
        END_IF;
        normalMode := FALSE;
    ELSE
        normalMode := TRUE;
        eT := tempSP - tempPV;
        eF := flowSP - flowPV;
        IF mode = 2 THEN
            trialT := accT + 0.2 * eT * scanSeconds;
            flowSPLimit := LIMIT(0.0, 1.0 * eT + trialT, 50.0);
            flowSP := flowSPLimit;
            accT := flowSP - 1.0 * eT;
            eF := flowSP - flowPV;
            trialF := accF + 0.5 * eF * scanSeconds;
            valveLimit := LIMIT(0.0, 2.0 * eF + trialF, 100.0);
            valveCommand := valveLimit;
            accF := valveCommand - 2.0 * eF;
        ELSIF mode = 1 THEN
            flowSP := manualFlowSP;
            eF := flowSP - flowPV;
            trialF := accF + 0.5 * eF * scanSeconds;
            valveLimit := LIMIT(0.0, 2.0 * eF + trialF, 100.0);
            valveCommand := valveLimit;
            accF := valveCommand - 2.0 * eF;
        ELSE
            flowSP := manualFlowSP;
            valveCommand := manualValve;
            accF := valveCommand - 2.0 * eF;
        END_IF;
    END_IF;

    prevResetBtn := resetBtn;
    prevMode := mode;
    prevFlowSP := flowSP;
    prevValveCommand := valveCommand;
    firstScanDone := TRUE;
END_FUNCTION_BLOCK

(* ---- self-medium-01.candidate_01.st ---- *)
FUNCTION_BLOCK FB
VAR_INPUT
    recipe   : ARRAY[1..8] OF ST_Recipe;
    selSlot  : INT;
    loadCmd  : BOOL;
    running  : BOOL;
END_VAR

VAR_OUTPUT
    valid    : BOOL;
    loadedID : INT;
END_VAR

VAR
    prevLoadCmd : BOOL := FALSE;
    prevRunning : BOOL := FALSE;
    prevValid   : BOOL := FALSE;
    prevLoadedID: INT  := 0;
END_VAR

VAR_TEMP
    risingEdge : BOOL;
    slotValid  : BOOL;
END_VAR

// Detect rising edge of loadCmd
risingEdge := loadCmd AND NOT prevLoadCmd;

// State retention: hold previous values unless explicitly updated
valid   := prevValid;
loadedID := prevLoadedID;

// Process load command only on rising edge and when not running
IF risingEdge AND NOT running THEN
    // Bounds check before array access
    IF (selSlot >= 1) AND (selSlot <= 8) THEN
        // Check all three validation conditions
        slotValid := (recipe[selSlot].recipeID <> 0)
                     AND (recipe[selSlot].totalRatio >= 99.0)
                     AND (recipe[selSlot].totalRatio <= 101.0)
                     AND (recipe[selSlot].temperature >= 30.0)
                     AND (recipe[selSlot].temperature <= 180.0);

        valid    := slotValid;
        loadedID := 0; // default on invalid
        IF slotValid THEN
            loadedID := recipe[selSlot].recipeID;
        END_IF;
    ELSE
        // Out-of-bounds: mark invalid, do not access array
        valid    := FALSE;
        loadedID := 0;
    END_IF;
END_IF;

// Update previous-cycle state for next scan
prevLoadCmd  := loadCmd;
prevRunning  := running;
prevValid    := valid;
prevLoadedID := loadedID;

END_FUNCTION_BLOCK

(* ---- self-medium-01.candidate_02.st ---- *)
TYPE ST_Recipe : STRUCT
    recipeID    : INT;
    totalRatio  : REAL;
    temperature : REAL;
END_STRUCT;
END_TYPE;

FUNCTION_BLOCK FB
VAR_INPUT
    recipe   : ARRAY[1..8] OF ST_Recipe;
    selSlot  : INT;
    loadCmd  : BOOL;
    running  : BOOL;
END_VAR

VAR_OUTPUT
    valid    : BOOL;
    loadedID : INT;
END_VAR

VAR
    prevLoadCmd  : BOOL := FALSE;
    prevRunning  : BOOL := FALSE;
    prevValid    : BOOL := FALSE;
    prevLoadedID : INT  := 0;
END_VAR

VAR_TEMP
    curRecipeID  : INT;
    curRatio     : REAL;
    curTemp      : REAL;
    slotInBounds : BOOL;
    recipeNotEmpty : BOOL;
    ratioInRange : BOOL;
    tempInRange  : BOOL;
    loadValid    : BOOL;
END_VAR

// Default: retain previous state
valid    := prevValid;
loadedID := prevLoadedID;

// Rising edge detection of loadCmd
IF loadCmd AND NOT prevLoadCmd THEN
    // Only process when not running
    IF NOT running THEN
        // Bounds check before array access
        slotInBounds := (selSlot >= 1) AND (selSlot <= 8);

        IF slotInBounds THEN
            // Read values into temporaries
            curRecipeID := recipe[selSlot].recipeID;
            curRatio    := recipe[selSlot].totalRatio;
            curTemp     := recipe[selSlot].temperature;

            // Validate each condition
            recipeNotEmpty := (curRecipeID <> 0);
            ratioInRange   := (curRatio >= 99.0) AND (curRatio <= 101.0);
            tempInRange    := (curTemp >= 30.0) AND (curTemp <= 180.0);

            // Combined validation
            loadValid := recipeNotEmpty AND ratioInRange AND tempInRange;

            valid    := loadValid;
            IF loadValid THEN
                loadedID := curRecipeID;
            ELSE
                loadedID := 0;
            END_IF;
        ELSE
            // Out-of-bounds: invalid, no array access
            valid    := FALSE;
            loadedID := 0;
        END_IF;
    END_IF;
END_IF;

// Update previous-cycle state
prevLoadCmd  := loadCmd;
prevRunning  := running;
prevValid    := valid;
prevLoadedID := loadedID;

END_FUNCTION_BLOCK

(* ---- self-medium-01.raw_candidate_01.st ---- *)
FUNCTION_BLOCK FB
VAR_INPUT
    recipe   : ARRAY[1..8] OF ST_Recipe;
    selSlot  : INT;
    loadCmd  : BOOL;
    running  : BOOL;
END_VAR

VAR_OUTPUT
    valid    : BOOL;
    loadedID : INT;
END_VAR

VAR
    prevLoadCmd : BOOL := FALSE;
    prevRunning : BOOL := FALSE;
    prevValid   : BOOL := FALSE;
    prevLoadedID: INT  := 0;
END_VAR

VAR_TEMP
    risingEdge : BOOL;
    slotValid  : BOOL;
END_VAR

// Detect rising edge of loadCmd
risingEdge := loadCmd AND NOT prevLoadCmd;

// State retention: hold previous values unless explicitly updated
valid   := prevValid;
loadedID := prevLoadedID;

// Process load command only on rising edge and when not running
IF risingEdge AND NOT running THEN
    // Bounds check before array access
    IF (selSlot >= 1) AND (selSlot <= 8) THEN
        // Check all three validation conditions
        slotValid := (recipe[selSlot].recipeID <> 0)
                     AND (recipe[selSlot].totalRatio >= 99.0)
                     AND (recipe[selSlot].totalRatio <= 101.0)
                     AND (recipe[selSlot].temperature >= 30.0)
                     AND (recipe[selSlot].temperature <= 180.0);

        valid    := slotValid;
        loadedID := 0; // default on invalid
        IF slotValid THEN
            loadedID := recipe[selSlot].recipeID;
        END_IF;
    ELSE
        // Out-of-bounds: mark invalid, do not access array
        valid    := FALSE;
        loadedID := 0;
    END_IF;
END_IF;

// Update previous-cycle state for next scan
prevLoadCmd  := loadCmd;
prevRunning  := running;
prevValid    := valid;
prevLoadedID := loadedID;

END_FUNCTION_BLOCK

(* ---- self-medium-01.raw_candidate_02.st ---- *)
TYPE ST_Recipe : STRUCT
    recipeID    : INT;
    totalRatio  : REAL;
    temperature : REAL;
END_STRUCT
END_TYPE

FUNCTION_BLOCK FB
VAR_INPUT
    recipe   : ARRAY[1..8] OF ST_Recipe;
    selSlot  : INT;
    loadCmd  : BOOL;
    running  : BOOL;
END_VAR

VAR_OUTPUT
    valid    : BOOL;
    loadedID : INT;
END_VAR

VAR
    prevLoadCmd  : BOOL := FALSE;
    prevRunning  : BOOL := FALSE;
    prevValid    : BOOL := FALSE;
    prevLoadedID : INT  := 0;
END_VAR

VAR_TEMP
    curRecipeID  : INT;
    curRatio     : REAL;
    curTemp      : REAL;
    slotInBounds : BOOL;
    recipeNotEmpty : BOOL;
    ratioInRange : BOOL;
    tempInRange  : BOOL;
    loadValid    : BOOL;
END_VAR

// Default: retain previous state
valid    := prevValid;
loadedID := prevLoadedID;

// Rising edge detection of loadCmd
IF loadCmd AND NOT prevLoadCmd THEN
    // Only process when not running
    IF NOT running THEN
        // Bounds check before array access
        slotInBounds := (selSlot >= 1) AND (selSlot <= 8);

        IF slotInBounds THEN
            // Read values into temporaries
            curRecipeID := recipe[selSlot].recipeID;
            curRatio    := recipe[selSlot].totalRatio;
            curTemp     := recipe[selSlot].temperature;

            // Validate each condition
            recipeNotEmpty := (curRecipeID <> 0);
            ratioInRange   := (curRatio >= 99.0) AND (curRatio <= 101.0);
            tempInRange    := (curTemp >= 30.0) AND (curTemp <= 180.0);

            // Combined validation
            loadValid := recipeNotEmpty AND ratioInRange AND tempInRange;

            valid    := loadValid;
            IF loadValid THEN
                loadedID := curRecipeID;
            ELSE
                loadedID := 0;
            END_IF;
        ELSE
            // Out-of-bounds: invalid, no array access
            valid    := FALSE;
            loadedID := 0;
        END_IF;
    END_IF;
END_IF;

// Update previous-cycle state
prevLoadCmd  := loadCmd;
prevRunning  := running;
prevValid    := valid;
prevLoadedID := loadedID;

END_FUNCTION_BLOCK

(* ---- self-medium-02.candidate_01.st ---- *)
FUNCTION_BLOCK FB
VAR
    buffer    : ARRAY[0..7] OF REAL;
    writeIndex : INT := 0;
END_VAR
VAR_OUTPUT
    filteredValue : REAL;
    windowFull    : BOOL;
    sampleCount   : INT;
END_VAR
VAR_INPUT
    enable   : BOOL;
    rawValue : REAL;
END_VAR

    IF enable THEN
        buffer[writeIndex] := rawValue;
        writeIndex := (writeIndex + 1) MOD 8;

        IF sampleCount < 8 THEN
            sampleCount := sampleCount + 1;
        END_IF;

        VAR i      : INT;
        VAR sum    : REAL;
        VAR idx    : INT;
        sum := 0.0;
        FOR i := 0 TO sampleCount - 1 DO
            idx    := (writeIndex - sampleCount + 8) MOD 8 + i;
            sum    := sum + buffer[idx];
        END_FOR;
        filteredValue := sum / INT_TO_REAL(sampleCount);

        windowFull := (sampleCount = 8);
    ELSE
        writeIndex := 0;
        sampleCount := 0;
        windowFull  := FALSE;
    END_IF;
END_FUNCTION_BLOCK

(* ---- self-medium-02.candidate_02.st ---- *)
FUNCTION_BLOCK FB
VAR
    buffer     : ARRAY[0..7] OF REAL;
    writeIndex : INT := 0;
    i          : INT;
    sum        : REAL;
END_VAR
VAR_OUTPUT
    filteredValue : REAL;
    windowFull    : BOOL;
    sampleCount   : INT;
END_VAR
VAR_INPUT
    enable   : BOOL;
    rawValue : REAL;
END_VAR

    IF enable THEN
        buffer[writeIndex] := rawValue;
        writeIndex := (writeIndex + 1) MOD 8;

        IF sampleCount < 8 THEN
            sampleCount := sampleCount + 1;
        END_IF;

        sum := 0.0;
        FOR i := 0 TO sampleCount - 1 DO
            IF writeIndex > i THEN
                sum := sum + buffer[writeIndex - i - 1];
            ELSE
                sum := sum + buffer[writeIndex - i - 1 + 8];
            END_IF;
        END_FOR;
        filteredValue := sum / INT_TO_REAL(sampleCount);

        windowFull := (sampleCount = 8);
    ELSE
        writeIndex := 0;
        sampleCount := 0;
        windowFull  := FALSE;
    END_IF;
END_FUNCTION_BLOCK

(* ---- self-medium-02.raw_candidate_01.st ---- *)
FUNCTION_BLOCK FB
VAR
    buffer    : ARRAY[0..7] OF REAL;
    writeIndex : INT := 0;
END_VAR
VAR_OUTPUT
    filteredValue : REAL;
    windowFull    : BOOL;
    sampleCount   : INT;
END_VAR
VAR_INPUT
    enable   : BOOL;
    rawValue : REAL;
END_VAR

    IF enable THEN
        buffer[writeIndex] := rawValue;
        writeIndex := (writeIndex + 1) MOD 8;

        IF sampleCount < 8 THEN
            sampleCount := sampleCount + 1;
        END_IF;

        VAR i      : INT;
        VAR sum    : REAL;
        VAR idx    : INT;
        sum := 0.0;
        FOR i := 0 TO sampleCount - 1 DO
            idx    := (writeIndex - sampleCount + 8) MOD 8 + i;
            sum    := sum + buffer[idx];
        END_FOR;
        filteredValue := sum / INT_TO_REAL(sampleCount);

        windowFull := (sampleCount = 8);
    ELSE
        writeIndex := 0;
        sampleCount := 0;
        windowFull  := FALSE;
    END_IF;
END_FUNCTION_BLOCK

(* ---- self-medium-02.raw_candidate_02.st ---- *)
FUNCTION_BLOCK FB
VAR
    buffer     : ARRAY[0..7] OF REAL;
    writeIndex : INT := 0;
    i          : INT;
    sum        : REAL;
END_VAR
VAR_OUTPUT
    filteredValue : REAL;
    windowFull    : BOOL;
    sampleCount   : INT;
END_VAR
VAR_INPUT
    enable   : BOOL;
    rawValue : REAL;
END_VAR

    IF enable THEN
        buffer[writeIndex] := rawValue;
        writeIndex := (writeIndex + 1) MOD 8;

        IF sampleCount < 8 THEN
            sampleCount := sampleCount + 1;
        END_IF;

        sum := 0.0;
        FOR i := 0 TO sampleCount - 1 DO
            IF writeIndex > i THEN
                sum := sum + buffer[writeIndex - i - 1];
            ELSE
                sum := sum + buffer[writeIndex - i - 1 + 8];
            END_IF;
        END_FOR;
        filteredValue := sum / INT_TO_REAL(sampleCount);

        windowFull := (sampleCount = 8);
    ELSE
        writeIndex := 0;
        sampleCount := 0;
        windowFull  := FALSE;
    END_IF;
END_FUNCTION_BLOCK

(* ---- self-medium-03.candidate_01.st ---- *)
FUNCTION_BLOCK FB
VAR_INPUT
    openBtn    : BOOL;
    closeBtn   : BOOL;
    openLimit  : BOOL;
    closeLimit : BOOL;
    obstacle   : BOOL;
END_VAR
VAR_OUTPUT
    motorUp    : BOOL;
    motorDown  : BOOL;
    errorFlag  : BOOL;
END_VAR
VAR
    state        : INT;
    prevOpenBtn  : BOOL;
    prevCloseBtn : BOOL;
    prevObstacle : BOOL;
    prevMotorUp  : BOOL;
    prevMotorDown: BOOL;
    prevErrorFlag: BOOL;
END_VAR
VAR_CONSTANT
    IDLE    : INT := 0;
    OPENING : INT := 1;
    CLOSING : INT := 2;
    FAULT   : INT := 3;
END_VAR

    // Rising edge detection
    VAR
        openRising   : BOOL;
        closeRising  : BOOL;
        doubleRising : BOOL;
    END_VAR
    openRising   := openBtn AND NOT prevOpenBtn;
    closeRising  := closeBtn AND NOT prevCloseBtn;
    doubleRising := (openBtn AND closeBtn) AND NOT (prevOpenBtn AND prevCloseBtn);

    // State transitions
    CASE state OF
    IDLE:
        // Clear fault on double-button rising edge when no obstacle
        IF doubleRising AND NOT obstacle THEN
            errorFlag := FALSE;
        END_IF;

        // Start opening: new rising edge on openBtn, closeBtn not held, no open limit
        IF openRising AND NOT closeBtn AND NOT openLimit AND NOT errorFlag THEN
            state    := OPENING;
            motorUp  := TRUE;
            motorDown:= FALSE;
        // Start closing: new rising edge on closeBtn, openBtn not held, no close limit
        ELSIF closeRising AND NOT openBtn AND NOT closeLimit AND NOT errorFlag THEN
            state    := CLOSING;
            motorUp  := FALSE;
            motorDown:= TRUE;
        ELSE
            motorUp  := FALSE;
            motorDown:= FALSE;
        END_IF;

    OPENING:
        // Obstacle detected: enter FAULT immediately
        IF obstacle THEN
            state     := FAULT;
            errorFlag := TRUE;
            motorUp   := FALSE;
            motorDown := FALSE;
        // Open limit reached: stop and return to IDLE
        ELSIF openLimit THEN
            state     := IDLE;
            motorUp   := FALSE;
            motorDown := FALSE;
        ELSE
            motorUp   := TRUE;
            motorDown := FALSE;
        END_IF;

    CLOSING:
        // Obstacle detected: enter FAULT immediately
        IF obstacle THEN
            state     := FAULT;
            errorFlag := TRUE;
            motorUp   := FALSE;
            motorDown := FALSE;
        // Close limit reached: stop and return to IDLE
        ELSIF closeLimit THEN
            state     := IDLE;
            motorUp   := FALSE;
            motorDown := FALSE;
        ELSE
            motorUp   := FALSE;
            motorDown := TRUE;
        END_IF;

    FAULT:
        // Latched: stay in FAULT unless double-button rising edge appears with no obstacle
        IF prevErrorFlag AND NOT obstacle AND doubleRising THEN
            state     := IDLE;
            errorFlag := FALSE;
            motorUp   := FALSE;
            motorDown := FALSE;
        ELSE
            errorFlag := TRUE;
            motorUp   := FALSE;
            motorDown := FALSE;
        END_IF;
    END_CASE;

    // Latch error flag once set (overrides any later state logic)
    IF errorFlag THEN
        motorUp   := FALSE;
        motorDown := FALSE;
    END_IF;

    // Update previous-cycle state for next scan
    prevOpenBtn   := openBtn;
    prevCloseBtn  := closeBtn;
    prevObstacle  := obstacle;
    prevMotorUp   := motorUp;
    prevMotorDown := motorDown;
    prevErrorFlag := errorFlag;
END_FUNCTION_BLOCK

(* ---- self-medium-03.candidate_02.st ---- *)
FUNCTION_BLOCK FB
VAR_INPUT
    openBtn   : BOOL;
    closeBtn  : BOOL;
    openLimit : BOOL;
    closeLimit: BOOL;
    obstacle  : BOOL;
END_VAR
VAR_OUTPUT
    motorUp   : BOOL;
    motorDown : BOOL;
    errorFlag : BOOL;
END_VAR
VAR
    state        : INT;
    prevOpenBtn  : BOOL;
    prevCloseBtn : BOOL;
    prevObstacle : BOOL;
    prevErrorFlag: BOOL;
END_VAR

    // Sample inputs
    VAR
        openRising  : BOOL;
        closeRising : BOOL;
        bothRising  : BOOL;
    END_VAR
    openRising  := openBtn AND NOT prevOpenBtn;
    closeRising := closeBtn AND NOT prevCloseBtn;
    bothRising  := (openBtn AND closeBtn) AND NOT (prevOpenBtn AND prevCloseBtn);

    // Initialize outputs to off
    motorUp   := FALSE;
    motorDown := FALSE;

    // Obstacle handling has highest priority in all states
    IF obstacle THEN
        state     := 3; // FAULT
        errorFlag := TRUE;
        motorUp   := FALSE;
        motorDown := FALSE;
    ELSE
        CASE state OF
        0: // IDLE
            // Reset fault with dual-button rising edge while obstacle clear
            IF prevErrorFlag AND bothRising THEN
                errorFlag := FALSE;
                state    := 0;
            ELSE
                errorFlag := FALSE;
            END_IF;
            // Start opening: rising edge on openBtn, closeBtn not pressed, not at open limit
            IF openRising AND NOT closeBtn AND NOT openLimit THEN
                state    := 1; // OPENING
                motorUp  := TRUE;
            // Start closing: rising edge on closeBtn, openBtn not pressed, not at close limit
            ELSIF closeRising AND NOT openBtn AND NOT closeLimit THEN
                state    := 2; // CLOSING
                motorDown:= TRUE;
            END_IF;

        1: // OPENING
            // Stop when open limit reached
            IF openLimit THEN
                state  := 0;
            ELSE
                motorUp := TRUE;
            END_IF;

        2: // CLOSING
            // Stop when close limit reached
            IF closeLimit THEN
                state    := 0;
            ELSE
                motorDown := TRUE;
            END_IF;

        3: // FAULT
            errorFlag := TRUE;
            // Clear fault only when no obstacle and dual-button rising edge appears
            IF prevErrorFlag AND bothRising THEN
                state    := 0;
                errorFlag := FALSE;
            END_IF;
        END_CASE;
    END_IF;

    // Update previous-cycle samples
    prevOpenBtn   := openBtn;
    prevCloseBtn  := closeBtn;
    prevObstacle  := obstacle;
    prevErrorFlag := errorFlag;
END_FUNCTION_BLOCK

(* ---- self-medium-03.raw_candidate_01.st ---- *)
FUNCTION_BLOCK FB
VAR_INPUT
    openBtn    : BOOL;
    closeBtn   : BOOL;
    openLimit  : BOOL;
    closeLimit : BOOL;
    obstacle   : BOOL;
END_VAR
VAR_OUTPUT
    motorUp    : BOOL;
    motorDown  : BOOL;
    errorFlag  : BOOL;
END_VAR
VAR
    state        : INT;
    prevOpenBtn  : BOOL;
    prevCloseBtn : BOOL;
    prevObstacle : BOOL;
    prevMotorUp  : BOOL;
    prevMotorDown: BOOL;
    prevErrorFlag: BOOL;
END_VAR
VAR_CONSTANT
    IDLE    : INT := 0;
    OPENING : INT := 1;
    CLOSING : INT := 2;
    FAULT   : INT := 3;
END_VAR

    // Rising edge detection
    VAR
        openRising   : BOOL;
        closeRising  : BOOL;
        doubleRising : BOOL;
    END_VAR
    openRising   := openBtn AND NOT prevOpenBtn;
    closeRising  := closeBtn AND NOT prevCloseBtn;
    doubleRising := (openBtn AND closeBtn) AND NOT (prevOpenBtn AND prevCloseBtn);

    // State transitions
    CASE state OF
    IDLE:
        // Clear fault on double-button rising edge when no obstacle
        IF doubleRising AND NOT obstacle THEN
            errorFlag := FALSE;
        END_IF;

        // Start opening: new rising edge on openBtn, closeBtn not held, no open limit
        IF openRising AND NOT closeBtn AND NOT openLimit AND NOT errorFlag THEN
            state    := OPENING;
            motorUp  := TRUE;
            motorDown:= FALSE;
        // Start closing: new rising edge on closeBtn, openBtn not held, no close limit
        ELSIF closeRising AND NOT openBtn AND NOT closeLimit AND NOT errorFlag THEN
            state    := CLOSING;
            motorUp  := FALSE;
            motorDown:= TRUE;
        ELSE
            motorUp  := FALSE;
            motorDown:= FALSE;
        END_IF;

    OPENING:
        // Obstacle detected: enter FAULT immediately
        IF obstacle THEN
            state     := FAULT;
            errorFlag := TRUE;
            motorUp   := FALSE;
            motorDown := FALSE;
        // Open limit reached: stop and return to IDLE
        ELSIF openLimit THEN
            state     := IDLE;
            motorUp   := FALSE;
            motorDown := FALSE;
        ELSE
            motorUp   := TRUE;
            motorDown := FALSE;
        END_IF;

    CLOSING:
        // Obstacle detected: enter FAULT immediately
        IF obstacle THEN
            state     := FAULT;
            errorFlag := TRUE;
            motorUp   := FALSE;
            motorDown := FALSE;
        // Close limit reached: stop and return to IDLE
        ELSIF closeLimit THEN
            state     := IDLE;
            motorUp   := FALSE;
            motorDown := FALSE;
        ELSE
            motorUp   := FALSE;
            motorDown := TRUE;
        END_IF;

    FAULT:
        // Latched: stay in FAULT unless double-button rising edge appears with no obstacle
        IF prevErrorFlag AND NOT obstacle AND doubleRising THEN
            state     := IDLE;
            errorFlag := FALSE;
            motorUp   := FALSE;
            motorDown := FALSE;
        ELSE
            errorFlag := TRUE;
            motorUp   := FALSE;
            motorDown := FALSE;
        END_IF;
    END_CASE;

    // Latch error flag once set (overrides any later state logic)
    IF errorFlag THEN
        motorUp   := FALSE;
        motorDown := FALSE;
    END_IF;

    // Update previous-cycle state for next scan
    prevOpenBtn   := openBtn;
    prevCloseBtn  := closeBtn;
    prevObstacle  := obstacle;
    prevMotorUp   := motorUp;
    prevMotorDown := motorDown;
    prevErrorFlag := errorFlag;
END_FUNCTION_BLOCK

(* ---- self-medium-03.raw_candidate_02.st ---- *)
FUNCTION_BLOCK FB
VAR_INPUT
    openBtn   : BOOL;
    closeBtn  : BOOL;
    openLimit : BOOL;
    closeLimit: BOOL;
    obstacle  : BOOL;
END_VAR
VAR_OUTPUT
    motorUp   : BOOL;
    motorDown : BOOL;
    errorFlag : BOOL;
END_VAR
VAR
    state        : INT;
    prevOpenBtn  : BOOL;
    prevCloseBtn : BOOL;
    prevObstacle : BOOL;
    prevErrorFlag: BOOL;
END_VAR

    // Sample inputs
    VAR
        openRising  : BOOL;
        closeRising : BOOL;
        bothRising  : BOOL;
    END_VAR
    openRising  := openBtn AND NOT prevOpenBtn;
    closeRising := closeBtn AND NOT prevCloseBtn;
    bothRising  := (openBtn AND closeBtn) AND NOT (prevOpenBtn AND prevCloseBtn);

    // Initialize outputs to off
    motorUp   := FALSE;
    motorDown := FALSE;

    // Obstacle handling has highest priority in all states
    IF obstacle THEN
        state     := 3; // FAULT
        errorFlag := TRUE;
        motorUp   := FALSE;
        motorDown := FALSE;
    ELSE
        CASE state OF
        0: // IDLE
            // Reset fault with dual-button rising edge while obstacle clear
            IF prevErrorFlag AND bothRising THEN
                errorFlag := FALSE;
                state    := 0;
            ELSE
                errorFlag := FALSE;
            END_IF;
            // Start opening: rising edge on openBtn, closeBtn not pressed, not at open limit
            IF openRising AND NOT closeBtn AND NOT openLimit THEN
                state    := 1; // OPENING
                motorUp  := TRUE;
            // Start closing: rising edge on closeBtn, openBtn not pressed, not at close limit
            ELSIF closeRising AND NOT openBtn AND NOT closeLimit THEN
                state    := 2; // CLOSING
                motorDown:= TRUE;
            END_IF;

        1: // OPENING
            // Stop when open limit reached
            IF openLimit THEN
                state  := 0;
            ELSE
                motorUp := TRUE;
            END_IF;

        2: // CLOSING
            // Stop when close limit reached
            IF closeLimit THEN
                state    := 0;
            ELSE
                motorDown := TRUE;
            END_IF;

        3: // FAULT
            errorFlag := TRUE;
            // Clear fault only when no obstacle and dual-button rising edge appears
            IF prevErrorFlag AND bothRising THEN
                state    := 0;
                errorFlag := FALSE;
            END_IF;
        END_CASE;
    END_IF;

    // Update previous-cycle samples
    prevOpenBtn   := openBtn;
    prevCloseBtn  := closeBtn;
    prevObstacle  := obstacle;
    prevErrorFlag := errorFlag;
END_FUNCTION_BLOCK

(* ---- self-medium-04.candidate_01.st ---- *)
FUNCTION_BLOCK FB
VAR_INPUT
    startBtn    : BOOL;
    resetBtn    : BOOL;
    doneSensor  : BOOL;
    targetVol   : REAL;
    flowVol     : REAL;
END_VAR
VAR_OUTPUT
    valveOpen   : BOOL;
    fillsToday  : INT;
END_VAR
VAR
    prevStartBtn      : BOOL := FALSE;
    prevResetBtn      : BOOL := FALSE;
    prevValveOpen     : BOOL := FALSE;
    currentVolume     : REAL := 0.0;
    pendingConfirm    : BOOL := FALSE;
    prevFillsToday    : INT  := 0;
END_VAR
VAR_TEMP
    risingStart  : BOOL;
    risingReset  : BOOL;
END_VAR
BEGIN
    risingStart  := startBtn AND NOT prevStartBtn;
    risingReset  := resetBtn AND NOT prevResetBtn;

    // Reset takes absolute priority
    IF risingReset THEN
        valveOpen      := FALSE;
        currentVolume  := 0.0;
        pendingConfirm := FALSE;
        fillsToday     := 0;
        prevFillsToday := 0;
    ELSIF risingStart THEN
        // New bottle starts
        pendingConfirm := FALSE;
        currentVolume  := flowVol;
        IF prevValveOpen THEN
            // Previous bottle still filling; cancel it, start new one
            valveOpen := TRUE;
        ELSE
            // Normal start from idle
            valveOpen := TRUE;
        END_IF;
        // Self-resetting: if this single shot already meets target
        IF currentVolume >= targetVol THEN
            valveOpen := FALSE;
            IF doneSensor THEN
                // Immediate confirmation same scan
                IF fillsToday < INT#32767 THEN
                    fillsToday := fillsToday + INT#1;
                END_IF;
                pendingConfirm := FALSE;
            ELSE
                pendingConfirm := TRUE;
            END_IF;
        END_IF;
    ELSIF valveOpen THEN
        // Currently filling: accumulate flow
        currentVolume := currentVolume + flowVol;
        IF currentVolume >= targetVol THEN
            valveOpen := FALSE;
            IF doneSensor THEN
                // Target met and sensor already true → confirm immediately
                IF fillsToday < INT#32767 THEN
                    fillsToday := fillsToday + INT#1;
                END_IF;
                pendingConfirm := FALSE;
            ELSE
                pendingConfirm := TRUE;
            END_IF;
        END_IF;
    ELSIF pendingConfirm THEN
        // Waiting for sensor confirmation
        valveOpen := FALSE;
        IF doneSensor THEN
            IF fillsToday < INT#32767 THEN
                fillsToday := fillsToday + INT#1;
            END_IF;
            pendingConfirm := FALSE;
        END_IF;
    ELSE
        // Idle, nothing pending
        valveOpen := FALSE;
    END_IF;

    // Update edge detectors for next scan
    prevStartBtn  := startBtn;
    prevResetBtn  := resetBtn;
    prevValveOpen := valveOpen;
    prevFillsToday := fillsToday;
END_FUNCTION_BLOCK

(* ---- self-medium-04.candidate_02.st ---- *)
FUNCTION_BLOCK FB
VAR_INPUT
    startBtn    : BOOL;
    resetBtn    : BOOL;
    doneSensor  : BOOL;
    targetVol   : REAL;
    flowVol     : REAL;
END_VAR
VAR_OUTPUT
    valveOpen   : BOOL;
    fillsToday  : INT;
END_VAR
VAR
    prevStartBtn    : BOOL := FALSE;
    prevResetBtn    : BOOL := FALSE;
    prevValveOpen   : BOOL := FALSE;
    prevFillsToday  : INT  := 0;
    currentVolume   : REAL := 0.0;
    pendingConfirm  : BOOL := FALSE;
END_VAR
BEGIN
    // Reset takes absolute priority
    IF resetBtn AND NOT prevResetBtn THEN
        valveOpen      := FALSE;
        currentVolume  := 0.0;
        pendingConfirm := FALSE;
        fillsToday     := 0;
        prevFillsToday := 0;
    ELSIF startBtn AND NOT prevStartBtn THEN
        // New bottle starts
        pendingConfirm := FALSE;
        currentVolume  := flowVol;
        valveOpen      := TRUE;
        // Self-resetting: if this single shot already meets target
        IF currentVolume >= targetVol THEN
            valveOpen      := FALSE;
            pendingConfirm := FALSE;
            IF doneSensor THEN
                IF fillsToday < INT#32767 THEN
                    fillsToday := fillsToday + INT#1;
                END_IF;
            ELSE
                pendingConfirm := TRUE;
            END_IF;
        END_IF;
    ELSIF valveOpen THEN
        // Currently filling: accumulate flow
        currentVolume := currentVolume + flowVol;
        IF currentVolume >= targetVol THEN
            valveOpen      := FALSE;
            pendingConfirm := FALSE;
            IF doneSensor THEN
                IF fillsToday < INT#32767 THEN
                    fillsToday := fillsToday + INT#1;
                END_IF;
            ELSE
                pendingConfirm := TRUE;
            END_IF;
        END_IF;
    ELSIF pendingConfirm THEN
        // Waiting for sensor confirmation
        valveOpen := FALSE;
        IF doneSensor THEN
            IF fillsToday < INT#32767 THEN
                fillsToday := fillsToday + INT#1;
            END_IF;
            pendingConfirm := FALSE;
        END_IF;
    ELSE
        // Idle, nothing pending
        valveOpen := FALSE;
    END_IF;

    // Update edge detectors for next scan
    prevStartBtn   := startBtn;
    prevResetBtn   := resetBtn;
    prevValveOpen  := valveOpen;
    prevFillsToday := fillsToday;
END_FUNCTION_BLOCK

(* ---- self-medium-04.raw_candidate_01.st ---- *)
FUNCTION_BLOCK FB
VAR_INPUT
    startBtn    : BOOL;
    resetBtn    : BOOL;
    doneSensor  : BOOL;
    targetVol   : REAL;
    flowVol     : REAL;
END_VAR
VAR_OUTPUT
    valveOpen   : BOOL;
    fillsToday  : INT;
END_VAR
VAR
    prevStartBtn      : BOOL := FALSE;
    prevResetBtn      : BOOL := FALSE;
    prevValveOpen     : BOOL := FALSE;
    currentVolume     : REAL := 0.0;
    pendingConfirm    : BOOL := FALSE;
    prevFillsToday    : INT  := 0;
END_VAR
VAR_TEMP
    risingStart  : BOOL;
    risingReset  : BOOL;
END_VAR
BEGIN
    risingStart  := startBtn AND NOT prevStartBtn;
    risingReset  := resetBtn AND NOT prevResetBtn;

    // Reset takes absolute priority
    IF risingReset THEN
        valveOpen      := FALSE;
        currentVolume  := 0.0;
        pendingConfirm := FALSE;
        fillsToday     := 0;
        prevFillsToday := 0;
    ELSIF risingStart THEN
        // New bottle starts
        pendingConfirm := FALSE;
        currentVolume  := flowVol;
        IF prevValveOpen THEN
            // Previous bottle still filling; cancel it, start new one
            valveOpen := TRUE;
        ELSE
            // Normal start from idle
            valveOpen := TRUE;
        END_IF;
        // Self-resetting: if this single shot already meets target
        IF currentVolume >= targetVol THEN
            valveOpen := FALSE;
            IF doneSensor THEN
                // Immediate confirmation same scan
                IF fillsToday < INT#32767 THEN
                    fillsToday := fillsToday + INT#1;
                END_IF;
                pendingConfirm := FALSE;
            ELSE
                pendingConfirm := TRUE;
            END_IF;
        END_IF;
    ELSIF valveOpen THEN
        // Currently filling: accumulate flow
        currentVolume := currentVolume + flowVol;
        IF currentVolume >= targetVol THEN
            valveOpen := FALSE;
            IF doneSensor THEN
                // Target met and sensor already true → confirm immediately
                IF fillsToday < INT#32767 THEN
                    fillsToday := fillsToday + INT#1;
                END_IF;
                pendingConfirm := FALSE;
            ELSE
                pendingConfirm := TRUE;
            END_IF;
        END_IF;
    ELSIF pendingConfirm THEN
        // Waiting for sensor confirmation
        valveOpen := FALSE;
        IF doneSensor THEN
            IF fillsToday < INT#32767 THEN
                fillsToday := fillsToday + INT#1;
            END_IF;
            pendingConfirm := FALSE;
        END_IF;
    ELSE
        // Idle, nothing pending
        valveOpen := FALSE;
    END_IF;

    // Update edge detectors for next scan
    prevStartBtn  := startBtn;
    prevResetBtn  := resetBtn;
    prevValveOpen := valveOpen;
    prevFillsToday := fillsToday;
END_FUNCTION_BLOCK

(* ---- self-medium-04.raw_candidate_02.st ---- *)
FUNCTION_BLOCK FB
VAR_INPUT
    startBtn    : BOOL;
    resetBtn    : BOOL;
    doneSensor  : BOOL;
    targetVol   : REAL;
    flowVol     : REAL;
END_VAR
VAR_OUTPUT
    valveOpen   : BOOL;
    fillsToday  : INT;
END_VAR
VAR
    prevStartBtn    : BOOL := FALSE;
    prevResetBtn    : BOOL := FALSE;
    prevValveOpen   : BOOL := FALSE;
    prevFillsToday  : INT  := 0;
    currentVolume   : REAL := 0.0;
    pendingConfirm  : BOOL := FALSE;
END_VAR
BEGIN
    // Reset takes absolute priority
    IF resetBtn AND NOT prevResetBtn THEN
        valveOpen      := FALSE;
        currentVolume  := 0.0;
        pendingConfirm := FALSE;
        fillsToday     := 0;
        prevFillsToday := 0;
    ELSIF startBtn AND NOT prevStartBtn THEN
        // New bottle starts
        pendingConfirm := FALSE;
        currentVolume  := flowVol;
        valveOpen      := TRUE;
        // Self-resetting: if this single shot already meets target
        IF currentVolume >= targetVol THEN
            valveOpen      := FALSE;
            pendingConfirm := FALSE;
            IF doneSensor THEN
                IF fillsToday < INT#32767 THEN
                    fillsToday := fillsToday + INT#1;
                END_IF;
            ELSE
                pendingConfirm := TRUE;
            END_IF;
        END_IF;
    ELSIF valveOpen THEN
        // Currently filling: accumulate flow
        currentVolume := currentVolume + flowVol;
        IF currentVolume >= targetVol THEN
            valveOpen      := FALSE;
            pendingConfirm := FALSE;
            IF doneSensor THEN
                IF fillsToday < INT#32767 THEN
                    fillsToday := fillsToday + INT#1;
                END_IF;
            ELSE
                pendingConfirm := TRUE;
            END_IF;
        END_IF;
    ELSIF pendingConfirm THEN
        // Waiting for sensor confirmation
        valveOpen := FALSE;
        IF doneSensor THEN
            IF fillsToday < INT#32767 THEN
                fillsToday := fillsToday + INT#1;
            END_IF;
            pendingConfirm := FALSE;
        END_IF;
    ELSE
        // Idle, nothing pending
        valveOpen := FALSE;
    END_IF;

    // Update edge detectors for next scan
    prevStartBtn   := startBtn;
    prevResetBtn   := resetBtn;
    prevValveOpen  := valveOpen;
    prevFillsToday := fillsToday;
END_FUNCTION_BLOCK

(* ---- self-medium-05.candidate_01.st ---- *)
FUNCTION_BLOCK FB
VAR_INPUT
    enable        : BOOL;
    resetBtn      : BOOL;
    scanSeconds   : LREAL;
    steamFlow     : LREAL;
    fuelFlow      : LREAL;
    steamTemp     : LREAL;
    steamPressure : LREAL;
END_VAR

VAR_OUTPUT
    qualified    : BOOL;
    dataFault    : BOOL;
    qualifiedTon : LREAL;
    fuelTon      : LREAL;
    revenue      : LREAL;
    cost         : LREAL;
    netProfit    : LREAL;
END_VAR

VAR
    prevResetBtn     : BOOL := FALSE;
    prevQualifiedTon : LREAL := 0.0;
    prevFuelTon      : LREAL := 0.0;
END_VAR

// Determine qualified status (closed interval)
qualified := (steamTemp >= 447.0) AND (steamTemp <= 453.0) AND
             (steamPressure >= 3750.0) AND (steamPressure <= 3850.0);

// Determine data fault status
dataFault := (scanSeconds <= 0.0) OR (scanSeconds > 10.0) OR
             (steamFlow < 0.0) OR (steamFlow > 90.0) OR
             (fuelFlow < 0.0) OR (fuelFlow > 6.0);

// Store previous cycle values for formula verification
prevQualifiedTon := qualifiedTon;
prevFuelTon := fuelTon;

// Reset rising edge takes priority over fault freeze
IF resetBtn AND NOT prevResetBtn THEN
    qualifiedTon := 0.0;
    fuelTon := 0.0;
ELSIF enable AND NOT dataFault THEN
    qualifiedTon := qualifiedTon + steamFlow * scanSeconds / 1000.0;
    fuelTon := fuelTon + fuelFlow * scanSeconds / 1000.0;
ELSE
    qualifiedTon := qualifiedTon;
    fuelTon := fuelTon;
END_IF;

// Update previous reset state for next cycle edge detection
prevResetBtn := resetBtn;

// Revenue, cost, and net profit updated every scan
revenue := qualifiedTon * 280.0;
cost := fuelTon * 1500.0;
netProfit := revenue - cost;

END_FUNCTION_BLOCK

(* ---- self-medium-05.candidate_02.st ---- *)
FUNCTION_BLOCK FB
VAR_INPUT
    enable        : BOOL;
    resetBtn      : BOOL;
    scanSeconds   : LREAL;
    steamFlow     : LREAL;
    fuelFlow      : LREAL;
    steamTemp     : LREAL;
    steamPressure : LREAL;
END_VAR

VAR_OUTPUT
    qualified    : BOOL;
    dataFault    : BOOL;
    qualifiedTon : LREAL;
    fuelTon      : LREAL;
    revenue      : LREAL;
    cost         : LREAL;
    netProfit    : LREAL;
END_VAR

VAR
    prevResetBtn : BOOL := FALSE;
END_VAR

// Data fault: scanSeconds not in (0,10] or flows out of range
dataFault := (scanSeconds <= 0.0) OR (scanSeconds > 10.0) OR
             (steamFlow < 0.0) OR (steamFlow > 90.0) OR
             (fuelFlow < 0.0) OR (fuelFlow > 6.0);

// Qualified: steamTemp in [446,453] AND steamPressure in [3750,3850]
qualified := (steamTemp >= 446.0) AND (steamTemp <= 453.0) AND
             (steamPressure >= 3750.0) AND (steamPressure <= 3850.0);

// Reset rising edge takes priority - clear and skip accumulation
IF resetBtn AND NOT prevResetBtn THEN
    qualifiedTon := 0.0;
    fuelTon := 0.0;
ELSIF enable AND NOT dataFault THEN
    // Fuel accumulates whenever enabled and no fault
    fuelTon := fuelTon + fuelFlow * scanSeconds / 1000.0;
    // Qualified steam accumulates only when qualified
    IF qualified THEN
        qualifiedTon := qualifiedTon + steamFlow * scanSeconds / 1000.0;
    END_IF;
END_IF;

// Store reset state for edge detection
prevResetBtn := resetBtn;

// Revenue, cost, netProfit updated every scan
revenue := qualifiedTon * 280.0;
cost := fuelTon * 1500.0;
netProfit := revenue - cost;

END_FUNCTION_BLOCK

(* ---- self-medium-05.raw_candidate_01.st ---- *)
FUNCTION_BLOCK FB
VAR_INPUT
    enable        : BOOL;
    resetBtn      : BOOL;
    scanSeconds   : LREAL;
    steamFlow     : LREAL;
    fuelFlow      : LREAL;
    steamTemp     : LREAL;
    steamPressure : LREAL;
END_VAR

VAR_OUTPUT
    qualified    : BOOL;
    dataFault    : BOOL;
    qualifiedTon : LREAL;
    fuelTon      : LREAL;
    revenue      : LREAL;
    cost         : LREAL;
    netProfit    : LREAL;
END_VAR

VAR
    prevResetBtn     : BOOL := FALSE;
    prevQualifiedTon : LREAL := 0.0;
    prevFuelTon      : LREAL := 0.0;
END_VAR

// Determine qualified status (closed interval)
qualified := (steamTemp >= 447.0) AND (steamTemp <= 453.0) AND
             (steamPressure >= 3750.0) AND (steamPressure <= 3850.0);

// Determine data fault status
dataFault := (scanSeconds <= 0.0) OR (scanSeconds > 10.0) OR
             (steamFlow < 0.0) OR (steamFlow > 90.0) OR
             (fuelFlow < 0.0) OR (fuelFlow > 6.0);

// Store previous cycle values for formula verification
prevQualifiedTon := qualifiedTon;
prevFuelTon := fuelTon;

// Reset rising edge takes priority over fault freeze
IF resetBtn AND NOT prevResetBtn THEN
    qualifiedTon := 0.0;
    fuelTon := 0.0;
ELSIF enable AND NOT dataFault THEN
    qualifiedTon := qualifiedTon + steamFlow * scanSeconds / 1000.0;
    fuelTon := fuelTon + fuelFlow * scanSeconds / 1000.0;
ELSE
    qualifiedTon := qualifiedTon;
    fuelTon := fuelTon;
END_IF;

// Update previous reset state for next cycle edge detection
prevResetBtn := resetBtn;

// Revenue, cost, and net profit updated every scan
revenue := qualifiedTon * 280.0;
cost := fuelTon * 1500.0;
netProfit := revenue - cost;

END_FUNCTION_BLOCK

(* ---- self-medium-05.raw_candidate_02.st ---- *)
FUNCTION_BLOCK FB
VAR_INPUT
    enable        : BOOL;
    resetBtn      : BOOL;
    scanSeconds   : LREAL;
    steamFlow     : LREAL;
    fuelFlow      : LREAL;
    steamTemp     : LREAL;
    steamPressure : LREAL;
END_VAR

VAR_OUTPUT
    qualified    : BOOL;
    dataFault    : BOOL;
    qualifiedTon : LREAL;
    fuelTon      : LREAL;
    revenue      : LREAL;
    cost         : LREAL;
    netProfit    : LREAL;
END_VAR

VAR
    prevResetBtn : BOOL := FALSE;
END_VAR

// Data fault: scanSeconds not in (0,10] or flows out of range
dataFault := (scanSeconds <= 0.0) OR (scanSeconds > 10.0) OR
             (steamFlow < 0.0) OR (steamFlow > 90.0) OR
             (fuelFlow < 0.0) OR (fuelFlow > 6.0);

// Qualified: steamTemp in [446,453] AND steamPressure in [3750,3850]
qualified := (steamTemp >= 446.0) AND (steamTemp <= 453.0) AND
             (steamPressure >= 3750.0) AND (steamPressure <= 3850.0);

// Reset rising edge takes priority - clear and skip accumulation
IF resetBtn AND NOT prevResetBtn THEN
    qualifiedTon := 0.0;
    fuelTon := 0.0;
ELSIF enable AND NOT dataFault THEN
    // Fuel accumulates whenever enabled and no fault
    fuelTon := fuelTon + fuelFlow * scanSeconds / 1000.0;
    // Qualified steam accumulates only when qualified
    IF qualified THEN
        qualifiedTon := qualifiedTon + steamFlow * scanSeconds / 1000.0;
    END_IF;
END_IF;

// Store reset state for edge detection
prevResetBtn := resetBtn;

// Revenue, cost, netProfit updated every scan
revenue := qualifiedTon * 280.0;
cost := fuelTon * 1500.0;
netProfit := revenue - cost;

END_FUNCTION_BLOCK

(* ---- self-medium-06.candidate_01.st ---- *)
FUNCTION_BLOCK FB
VAR_INPUT
    enable         : BOOL;
    resetBtn       : BOOL;
    sensorValid    : BOOL;
    setpoint       : REAL;
    temperature    : REAL;
    scanSeconds    : REAL;
    bias           : REAL;
END_VAR
VAR_OUTPUT
    power          : REAL;
    correction     : REAL;
    fault          : BOOL;
END_VAR
VAR
    ePrev          : REAL := 0.0;
    historyFirst   : BOOL := FALSE;
    resetPrev      : BOOL := FALSE;
END_VAR
VAR_TEMP
    e              : REAL;
    de             : REAL;
    xNorm          : REAL;
    yNorm          : REAL;
    muNx           : REAL;
    muZx           : REAL;
    muPx           : REAL;
    muNy           : REAL;
    muZy           : REAL;
    muPy           : REAL;
    wNN            : REAL;
    wNZ            : REAL;
    wNP            : REAL;
    wZN            : REAL;
    wZZ            : REAL;
    wZP            : REAL;
    wPN            : REAL;
    wPZ            : REAL;
    wPP            : REAL;
    sumW           : REAL;
    sumWC          : REAL;
    risingReset    : BOOL;
    firstScan      : BOOL;
END_VAR
BEGIN
    risingReset := resetBtn AND NOT resetPrev;
    resetPrev   := resetBtn;

    fault := NOT sensorValid OR scanSeconds <= 0.0 OR scanSeconds > 10.0;

    IF NOT enable OR fault OR risingReset THEN
        power       := 0.0;
        correction  := 0.0;
        ePrev       := 0.0;
        historyFirst := FALSE;
    ELSE
        e := setpoint - temperature;

        IF NOT historyFirst THEN
            de := 0.0;
        ELSE
            de := (e - ePrev) / scanSeconds;
        END_IF;

        xNorm := LIMIT(-1.0, e / 10.0, 1.0);
        yNorm := LIMIT(-1.0, de / 2.0, 1.0);

        muNx := MAX(-xNorm, 0.0);
        muZx := MAX(1.0 - ABS(xNorm), 0.0);
        muPx := MAX(xNorm, 0.0);

        muNy := MAX(-yNorm, 0.0);
        muZy := MAX(1.0 - ABS(yNorm), 0.0);
        muPy := MAX(yNorm, 0.0);

        wNN := muNx * muNy;
        wNZ := muNx * muZy;
        wNP := muNx * muPy;
        wZN := muZx * muNy;
        wZZ := muZx * muZy;
        wZP := muZx * muPy;
        wPN := muPx * muNy;
        wPZ := muPx * muZy;
        wPP := muPx * muPy;

        sumW := wNN + wNZ + wNP + wZN + wZZ + wZP + wPN + wPZ + wPP;

        sumWC := wNN * (-30.0)
               + wNZ * (-20.0)
               + wNP * (-10.0)
               + wZN * (-10.0)
               + wZZ *   0.0
               + wZP *  10.0
               + wPN *  10.0
               + wPZ *  20.0
               + wPP *  30.0;

        IF sumW > 0.0 THEN
            correction := sumWC / sumW;
        ELSE
            correction := 0.0;
        END_IF;

        power := LIMIT(0.0, bias + correction, 100.0);

        firstScan := NOT historyFirst;
        ePrev := e;
        historyFirst := TRUE;
    END_IF;
END_FUNCTION_BLOCK

(* ---- self-medium-06.candidate_02.st ---- *)
FUNCTION_BLOCK FB
VAR_INPUT
    enable       : BOOL;
    resetBtn     : BOOL;
    sensorValid  : BOOL;
    setpoint     : REAL;
    temperature  : REAL;
    scanSeconds  : REAL;
    bias         : REAL;
END_VAR
VAR_OUTPUT
    power       : REAL;
    correction  : REAL;
    fault       : BOOL;
END_VAR
VAR
    ePrev        : REAL := 0.0;
    historyValid : BOOL := FALSE;
    prevReset    : BOOL := FALSE;
    e            : REAL;
    de           : REAL;
    xNorm        : REAL;
    yNorm        : REAL;
    muNx         : REAL;
    muZx         : REAL;
    muPx         : REAL;
    muNy         : REAL;
    muZy         : REAL;
    muPy         : REAL;
    wNN          : REAL;
    wNZ          : REAL;
    wNP          : REAL;
    wZN          : REAL;
    wZZ          : REAL;
    wZP          : REAL;
    wPN          : REAL;
    wPZ          : REAL;
    wPP          : REAL;
    sumW         : REAL;
    sumWC        : REAL;
END_VAR
BEGIN
    fault := NOT sensorValid OR scanSeconds <= 0.0 OR scanSeconds > 10.0;

    IF NOT enable OR fault OR (resetBtn AND NOT prevReset) THEN
        power      := 0.0;
        correction := 0.0;
        ePrev      := 0.0;
        historyValid := FALSE;
    ELSE
        e := setpoint - temperature;

        IF NOT historyValid THEN
            de := 0.0;
        ELSE
            de := (e - ePrev) / scanSeconds;
        END_IF;

        xNorm := LIMIT(-1.0, e / 10.0, 1.0);
        yNorm := LIMIT(-1.0, de / 2.0, 1.0);

        muNx := MAX(-xNorm, 0.0);
        muZx := MAX(1.0 - ABS(xNorm), 0.0);
        muPx := MAX(xNorm, 0.0);

        muNy := MAX(-yNorm, 0.0);
        muZy := MAX(1.0 - ABS(yNorm), 0.0);
        muPy := MAX(yNorm, 0.0);

        wNN := muNx * muNy;
        wNZ := muNx * muZy;
        wNP := muNx * muPy;
        wZN := muZx * muNy;
        wZZ := muZx * muZy;
        wZP := muZx * muPy;
        wPN := muPx * muNy;
        wPZ := muPx * muZy;
        wPP := muPx * muPy;

        sumW := wNN + wNZ + wNP + wZN + wZZ + wZP + wPN + wPZ + wPP;

        sumWC := wNN * (-30.0)
               + wNZ * (-20.0)
               + wNP * (-10.0)
               + wZN * (-10.0)
               + wZZ *   0.0
               + wZP *  10.0
               + wPN *  10.0
               + wPZ *  20.0
               + wPP *  30.0;

        IF sumW > 0.0 THEN
            correction := sumWC / sumW;
        ELSE
            correction := 0.0;
        END_IF;

        power := LIMIT(0.0, bias + correction, 100.0);

        ePrev := e;
        historyValid := TRUE;
    END_IF;

    prevReset := resetBtn;
END_FUNCTION_BLOCK

(* ---- self-medium-06.raw_candidate_01.st ---- *)
FUNCTION_BLOCK FB
VAR_INPUT
    enable         : BOOL;
    resetBtn       : BOOL;
    sensorValid    : BOOL;
    setpoint       : REAL;
    temperature    : REAL;
    scanSeconds    : REAL;
    bias           : REAL;
END_VAR
VAR_OUTPUT
    power          : REAL;
    correction     : REAL;
    fault          : BOOL;
END_VAR
VAR
    ePrev          : REAL := 0.0;
    historyFirst   : BOOL := FALSE;
    resetPrev      : BOOL := FALSE;
END_VAR
VAR_TEMP
    e              : REAL;
    de             : REAL;
    xNorm          : REAL;
    yNorm          : REAL;
    muNx           : REAL;
    muZx           : REAL;
    muPx           : REAL;
    muNy           : REAL;
    muZy           : REAL;
    muPy           : REAL;
    wNN            : REAL;
    wNZ            : REAL;
    wNP            : REAL;
    wZN            : REAL;
    wZZ            : REAL;
    wZP            : REAL;
    wPN            : REAL;
    wPZ            : REAL;
    wPP            : REAL;
    sumW           : REAL;
    sumWC          : REAL;
    risingReset    : BOOL;
    firstScan      : BOOL;
END_VAR
BEGIN
    risingReset := resetBtn AND NOT resetPrev;
    resetPrev   := resetBtn;

    fault := NOT sensorValid OR scanSeconds <= 0.0 OR scanSeconds > 10.0;

    IF NOT enable OR fault OR risingReset THEN
        power       := 0.0;
        correction  := 0.0;
        ePrev       := 0.0;
        historyFirst := FALSE;
    ELSE
        e := setpoint - temperature;

        IF NOT historyFirst THEN
            de := 0.0;
        ELSE
            de := (e - ePrev) / scanSeconds;
        END_IF;

        xNorm := LIMIT(-1.0, e / 10.0, 1.0);
        yNorm := LIMIT(-1.0, de / 2.0, 1.0);

        muNx := MAX(-xNorm, 0.0);
        muZx := MAX(1.0 - ABS(xNorm), 0.0);
        muPx := MAX(xNorm, 0.0);

        muNy := MAX(-yNorm, 0.0);
        muZy := MAX(1.0 - ABS(yNorm), 0.0);
        muPy := MAX(yNorm, 0.0);

        wNN := muNx * muNy;
        wNZ := muNx * muZy;
        wNP := muNx * muPy;
        wZN := muZx * muNy;
        wZZ := muZx * muZy;
        wZP := muZx * muPy;
        wPN := muPx * muNy;
        wPZ := muPx * muZy;
        wPP := muPx * muPy;

        sumW := wNN + wNZ + wNP + wZN + wZZ + wZP + wPN + wPZ + wPP;

        sumWC := wNN * (-30.0)
               + wNZ * (-20.0)
               + wNP * (-10.0)
               + wZN * (-10.0)
               + wZZ *   0.0
               + wZP *  10.0
               + wPN *  10.0
               + wPZ *  20.0
               + wPP *  30.0;

        IF sumW > 0.0 THEN
            correction := sumWC / sumW;
        ELSE
            correction := 0.0;
        END_IF;

        power := LIMIT(0.0, bias + correction, 100.0);

        firstScan := NOT historyFirst;
        ePrev := e;
        historyFirst := TRUE;
    END_IF;
END_FUNCTION_BLOCK

(* ---- self-medium-06.raw_candidate_02.st ---- *)
FUNCTION_BLOCK FB
VAR_INPUT
    enable       : BOOL;
    resetBtn     : BOOL;
    sensorValid  : BOOL;
    setpoint     : REAL;
    temperature  : REAL;
    scanSeconds  : REAL;
    bias         : REAL;
END_VAR
VAR_OUTPUT
    power       : REAL;
    correction  : REAL;
    fault       : BOOL;
END_VAR
VAR
    ePrev        : REAL := 0.0;
    historyValid : BOOL := FALSE;
    prevReset    : BOOL := FALSE;
    e            : REAL;
    de           : REAL;
    xNorm        : REAL;
    yNorm        : REAL;
    muNx         : REAL;
    muZx         : REAL;
    muPx         : REAL;
    muNy         : REAL;
    muZy         : REAL;
    muPy         : REAL;
    wNN          : REAL;
    wNZ          : REAL;
    wNP          : REAL;
    wZN          : REAL;
    wZZ          : REAL;
    wZP          : REAL;
    wPN          : REAL;
    wPZ          : REAL;
    wPP          : REAL;
    sumW         : REAL;
    sumWC        : REAL;
END_VAR
BEGIN
    fault := NOT sensorValid OR scanSeconds <= 0.0 OR scanSeconds > 10.0;

    IF NOT enable OR fault OR (resetBtn AND NOT prevReset) THEN
        power      := 0.0;
        correction := 0.0;
        ePrev      := 0.0;
        historyValid := FALSE;
    ELSE
        e := setpoint - temperature;

        IF NOT historyValid THEN
            de := 0.0;
        ELSE
            de := (e - ePrev) / scanSeconds;
        END_IF;

        xNorm := LIMIT(-1.0, e / 10.0, 1.0);
        yNorm := LIMIT(-1.0, de / 2.0, 1.0);

        muNx := MAX(-xNorm, 0.0);
        muZx := MAX(1.0 - ABS(xNorm), 0.0);
        muPx := MAX(xNorm, 0.0);

        muNy := MAX(-yNorm, 0.0);
        muZy := MAX(1.0 - ABS(yNorm), 0.0);
        muPy := MAX(yNorm, 0.0);

        wNN := muNx * muNy;
        wNZ := muNx * muZy;
        wNP := muNx * muPy;
        wZN := muZx * muNy;
        wZZ := muZx * muZy;
        wZP := muZx * muPy;
        wPN := muPx * muNy;
        wPZ := muPx * muZy;
        wPP := muPx * muPy;

        sumW := wNN + wNZ + wNP + wZN + wZZ + wZP + wPN + wPZ + wPP;

        sumWC := wNN * (-30.0)
               + wNZ * (-20.0)
               + wNP * (-10.0)
               + wZN * (-10.0)
               + wZZ *   0.0
               + wZP *  10.0
               + wPN *  10.0
               + wPZ *  20.0
               + wPP *  30.0;

        IF sumW > 0.0 THEN
            correction := sumWC / sumW;
        ELSE
            correction := 0.0;
        END_IF;

        power := LIMIT(0.0, bias + correction, 100.0);

        ePrev := e;
        historyValid := TRUE;
    END_IF;

    prevReset := resetBtn;
END_FUNCTION_BLOCK
